(* IEC 61131-3 sources: Industry-PLC-LLM/data/PLCBEAD_repo/PLCBEAD_PLCEmbed-main/PLC-BEAD/Source/PLC_Programs (part 15) *)

(* ---- INC.ST ---- *)
FUNCTION INC:INT
	VAR_INPUT
		X :	INT;
		D :	INT;
		M :	INT;
	END_VAR

	inc := (X + D + M + 1) MOD (M + 1);
END_FUNCTION

PROGRAM program0
  VAR
    LocalVar0 : INT;
	LocalVar1 : INT;
	LocalVar2 : INT;
	LocalOUT  : INT;
  END_VAR
  	LocalOUT := INC(LocalVar0, LocalVar1,LocalVar2);
END_PROGRAM

CONFIGURATION Config0
  RESOURCE Res0 ON PLC
    TASK task0(INTERVAL := T#20ms,PRIORITY := 0);
    PROGRAM instance0 WITH task0 : program0;
  END_RESOURCE
END_CONFIGURATION

(* ---- INC1.ST ---- *)
FUNCTION INC1:INT

	VAR_INPUT
		X :	INT;
		N :	INT;
	END_VAR

	IF X >= N - 1 THEN
		INC1 := 0;
	ELSE
		INC1 := X + 1;
	END_IF;
END_FUNCTION

PROGRAM program0
  VAR
	X :	INT;
	N :	INT;
    CEIL5_OUT : INT;
  END_VAR

  CEIL5_OUT := INC1(X, N);
END_PROGRAM

CONFIGURATION Config0

  RESOURCE Res0 ON PLC
    TASK task0(INTERVAL := T#20ms,PRIORITY := 0);
    PROGRAM instance0 WITH task0 : program0;
  END_RESOURCE
END_CONFIGURATION

(* ---- INC2.ST ---- *)
FUNCTION INC2:INT

	VAR_INPUT
		X :	INT;
		D :	INT;
		L :	INT;
		U :	INT;
	END_VAR

	VAR
		tmp :	INT;
	END_VAR

	tmp := U - L + 1;
	INC2 := (X + D - L + tmp) MOD tmp + L;

END_FUNCTION

PROGRAM program0
	VAR
		X :	INT;
		D :	INT;
		L :	INT;
		U :	INT;
		CEIL5_OUT : INT;
	END_VAR

  	CEIL5_OUT := INC2(X, D, L, U);
END_PROGRAM

CONFIGURATION Config0

	RESOURCE Res0 ON PLC
		TASK task0(INTERVAL := T#20ms,PRIORITY := 0);
		PROGRAM instance0 WITH task0 : program0;
	END_RESOURCE

END_CONFIGURATION

(* ---- INI_PARSER_BUF_DEMO.ST ---- *)
PROGRAM INI_PARSER_BUF_DEMO

	VAR

	END_VAR

	VAR_EXTERNAL

	END_VAR

	VAR
		SMTP_SERVER :	STRING;
		SMTP_FROM :	STRING;
		STATION_NAME :	STRING;
		STATION_IP :	STRING;
	END_VAR

	VAR
		IPB :	INI_PARSER_BUF;
		FS :	FILE_SERVER;
		FSD :	oscat_FILE_SERVER_DATA;
		PT :	oscat_NETWORK_BUFFER;
		section :	INT;
		key :	oscat_STRING250;
		value :	oscat_STRING250;
		str :	oscat_STRING250;
		step :	INT;
		result :	BYTE;
		offset :	UDINT;
		run :	BYTE;
		done :	BOOL;
	END_VAR

	CASE step OF

	00:	IF NOT done then
			FSD.FILENAME := 'config.ini';
			FSD.MODE := BYTE#1;
			FSD.OFFSET := UDINT#0;
			FSD.AUTO_CLOSE := T#0s;
			PT.SIZE := UINT#65535;
			step := 10;
		END_IF;

	10:	IF FSD.MODE = BYTE#0 THEN
			offset := UDINT#0;
			str := '';
			run := BYTE#3;
			step := 50;
		END_IF;

	50:	IF run = BYTE#0 THEN
			run := BYTE#3;

			IF result = BYTE#1 THEN
				IF EQ_STRING(key,'Station') THEN
					section := 1;
				ELSIF EQ_STRING(key,'SMTP') THEN
					section := 2;

				ELSE
					section := 0;
				END_IF;

			ELSIF result = BYTE#2 AND section > 0 THEN

				CASE section OF

				1:
					IF EQ_STRING(key,'NAME') THEN
						STATION_NAME := value;
					ELSIF EQ_STRING(key,'IP') THEN
						STATION_IP := value;
					END_IF;

				2:
					IF EQ_STRING(key,'SERVER') THEN
						SMTP_SERVER := value;
					ELSIF EQ_STRING(key,'FROM') THEN
						SMTP_FROM := value;
					END_IF;

				END_CASE;

			ELSIF result = BYTE#10 THEN
				run := BYTE#0;
				FSD.MODE := BYTE#5;
				step := 80;
			END_IF;
		END_IF;

	80:	IF FSD.MODE = BYTE#0 THEN
			done := TRUE;
			step := 0;
		END_IF;

	END_CASE;

	IPB(STR:=str,RUN:=run,OFFSET:=offset,KEY:=key,VALUE:=value,PT:=PT);
	str:=IPB.STR;
	run:=IPB.RUN;
	offset:=IPB.OFFSET;
	key:=IPB.KEY;
	value:=IPB.VALUE;
	PT:=IPB.PT;
	result:=IPB.RESULT;

	FS(FSD:=FSD,PT:=PT);
	FSD:=FS.FSD;
	PT:=FS.PT;

END_PROGRAM

(* ---- INI_PARSER_FILE_DEMO.ST ---- *)
PROGRAM INI_PARSER_FILE_DEMO

	VAR

	END_VAR

	VAR_EXTERNAL

	END_VAR

	VAR
		SMTP_SERVER :	STRING;
		SMTP_FROM :	STRING;
		STATION_NAME :	STRING;
		STATION_IP :	STRING;
	END_VAR

	VAR
		IPF :	INI_PARSER_FILE;
		FS :	FILE_SERVER;
		FSD :	oscat_FILE_SERVER_DATA;
		PT :	oscat_NETWORK_BUFFER;
		section :	INT;
		filename :	STRING;
		key :	oscat_STRING250;
		value :	oscat_STRING250;
		str :	oscat_STRING250;
		step :	INT;
		result :	BYTE;
		offset :	UDINT;
		run :	BYTE;
		done :	BOOL;
	END_VAR

	CASE step OF

	00:	IF NOT done THEN
			filename := 'config.ini';
			offset := UDINT#0;
			str := '';
			run := BYTE#3;
			step := 50;
		END_IF;

	50:	IF run = BYTE#0 THEN

			run := BYTE#3;

			IF result = BYTE#1 THEN
				IF EQ_STRING(key,'Station') THEN
					section := 1;
				ELSIF EQ_STRING(key,'SMTP') THEN
					section := 2;

				ELSE
					section := 0;
				END_IF;

			ELSIF result = BYTE#2 AND section > 0 THEN

				CASE section OF

				1:
					IF EQ_STRING(key,'NAME') THEN
						STATION_NAME := value;
					ELSIF EQ_STRING(key,'IP') THEN
						STATION_IP := value;
					END_IF;

				2:
					IF EQ_STRING(key,'SERVER') THEN
						SMTP_SERVER := value;
					ELSIF EQ_STRING(key,'FROM') THEN
						SMTP_FROM := value;
					END_IF;

				END_CASE;

			ELSIF result = BYTE#10 THEN
				run := BYTE#0;
				FSD.MODE := BYTE#5;
				step := 30;
			END_IF;
		END_IF;

	30:	IF FSD.MODE = BYTE#0 THEN
			step := 0;
			done := TRUE;
		END_IF;

	END_CASE;

	IPF(FILENAME:=FILENAME,FSD:=FSD,STR:=str,RUN:=run,OFFSET:=offset,KEY:=key,VALUE:=value,PT:=PT);
	FILENAME:=IPF.FILENAME;
	FSD:=IPF.FSD;
	str:=IPF.STR;
	run:=IPF.RUN;
	offset:=IPF.OFFSET;
	key:=IPF.KEY;
	value:=IPF.VALUE;
	PT:=IPF.PT;
	result:=IPF.RESULT;

	FS(FSD:=FSD,PT:=PT);
	FSD:=FS.FSD;
	PT:=FS.PT;

END_PROGRAM

(* ---- INT_TO_BCDC.ST ---- *)
FUNCTION INT_TO_BCDC:BYTE

	VAR_INPUT
		IN :	INT;
	END_VAR

	INT_TO_BCDC := SHL(INT_TO_BYTE(IN / INT#10),4) OR INT_TO_BYTE(in MOD INT#10);

END_FUNCTION

PROGRAM program0

	VAR
		IN :	INT;
		OUT : BYTE;
	END_VAR

	OUT := INT_TO_BCDC(IN);

END_PROGRAM

CONFIGURATION Config0

	RESOURCE Res0 ON PLC
		TASK task0(INTERVAL := T#20ms,PRIORITY := 0);
		PROGRAM instance0 WITH task0 : program0;
	END_RESOURCE

END_CONFIGURATION

(* ---- INT_TO_TIME.ST ---- *)
FUNCTION _INT_TO_TIME:TIME

	VAR_INPUT
		IN :	INT;
	END_VAR

	_INT_TO_TIME := DINT_TO_TIME(INT_TO_DINT(IN));

END_FUNCTION

PROGRAM program0
	VAR
		IN :	INT;
		OUT : TIME;
	END_VAR

	OUT := _INT_TO_TIME(IN);
END_PROGRAM

CONFIGURATION Config0

	RESOURCE Res0 ON PLC
		TASK task0(INTERVAL := T#20ms,PRIORITY := 0);
		PROGRAM instance0 WITH task0 : program0;
	END_RESOURCE

END_CONFIGURATION

(* ---- INV.ST ---- *)
FUNCTION INV:REAL

	VAR_INPUT
		X :	REAL;
	END_VAR

	IF X <> 0.0 THEN INV := 1.0 / X; END_IF;

END_FUNCTION

PROGRAM program0
	VAR
		X :	REAL;
		OUT : REAL;
	END_VAR

	OUT := INV(X);
END_PROGRAM

CONFIGURATION Config0

	RESOURCE Res0 ON PLC
		TASK task0(INTERVAL := T#20ms,PRIORITY := 0);
		PROGRAM instance0 WITH task0 : program0;
	END_RESOURCE

END_CONFIGURATION

(* ---- IP4_CHECK.ST ---- *)
FUNCTION IP4_CHECK:BOOL

	VAR_INPUT
		NIP :	DWORD;
		LIP :	DWORD;
		SM :	DWORD;
	END_VAR

	IP4_CHECK := (NIP AND sm) = (LIP AND SM);

END_FUNCTION

PROGRAM program0
	VAR
		NIP :	DWORD;
		LIP :	DWORD;
		SM :	DWORD;
		CEIL5_OUT : BOOL;
	END_VAR

  	CEIL5_OUT := IP4_CHECK(NIP, LIP, SM);
END_PROGRAM

CONFIGURATION Config0

  RESOURCE Res0 ON PLC
    TASK task0(INTERVAL := T#20ms,PRIORITY := 0);
    PROGRAM instance0 WITH task0 : program0;
  END_RESOURCE
END_CONFIGURATION

(* ---- IS_URLCHR.ST ---- *)
FUNCTION IS_URLCHR:BOOL

	VAR_INPUT
		IN :	BYTE;
	END_VAR

	IS_URLCHR := ((IN>BYTE#47) AND (IN<BYTE#58)) OR ((IN>BYTE#64) AND (IN<BYTE#91)) OR ((IN>BYTE#96) AND (IN<BYTE#123)) OR (in=BYTE#126) OR (in=BYTE#95) OR (in=BYTE#45) OR (in=BYTE#46);

END_FUNCTION

PROGRAM program0
	VAR
		IN :	BYTE;
		CEIL5_OUT : BOOL;
	END_VAR

  	CEIL5_OUT := IS_URLCHR(IN);
END_PROGRAM

CONFIGURATION Config0

  RESOURCE Res0 ON PLC
    TASK task0(INTERVAL := T#20ms,PRIORITY := 0);
    PROGRAM instance0 WITH task0 : program0;
  END_RESOURCE
END_CONFIGURATION

(* ---- ISC_ALPHA.ST ---- *)
FUNCTION SETUP_EXTENDED_ASCII:BOOL

	VAR_INPUT
		X :	BOOL;
	END_VAR

	SETUP_EXTENDED_ASCII := X OR TRUE;

END_FUNCTION

FUNCTION ISC_ALPHA:BOOL

	VAR_INPUT
		IN :	BYTE;
	END_VAR

	IF SETUP_EXTENDED_ASCII(FALSE) THEN
		ISC_ALPHA := (in > BYTE#64 AND in < BYTE#91) OR (in > BYTE#191  AND in <> BYTE#215 AND in <> BYTE#247) OR (in > BYTE#96 AND in < BYTE#123);
	ELSE
		ISC_ALPHA := (IN > BYTE#64 AND IN < BYTE#91) OR (in > BYTE#96 AND in < BYTE#123);
	END_IF;

END_FUNCTION

PROGRAM program0
	VAR
		IN : BYTE;
		OUT : BOOL;
	END_VAR

	OUT := ISC_ALPHA(IN);
END_PROGRAM

CONFIGURATION Config0

	RESOURCE Res0 ON PLC
		TASK task0(INTERVAL := T#20ms,PRIORITY := 0);
		PROGRAM instance0 WITH task0 : program0;
	END_RESOURCE

END_CONFIGURATION

(* ---- ISC_CTRL.ST ---- *)
FUNCTION ISC_CTRL:BOOL

	VAR_INPUT
		IN :	BYTE;
	END_VAR

	ISC_CTRL := IN < BYTE#32 OR IN = BYTE#127;

END_FUNCTION

PROGRAM program0
	VAR
		IN : BYTE;
		OUT : BOOL;
	END_VAR

	OUT := ISC_CTRL(IN);
END_PROGRAM

CONFIGURATION Config0

	RESOURCE Res0 ON PLC
		TASK task0(INTERVAL := T#20ms,PRIORITY := 0);
		PROGRAM instance0 WITH task0 : program0;
	END_RESOURCE

END_CONFIGURATION

(* ---- ISC_HEX.ST ---- *)
FUNCTION ISC_HEX:BOOL

	VAR_INPUT
		IN :	BYTE;
	END_VAR

	ISC_HEX := (IN > BYTE#47 AND IN < BYTE#58) OR (IN > BYTE#64 AND IN < BYTE#71) OR (IN > BYTE#96 AND IN < BYTE#103);

END_FUNCTION

PROGRAM program0
	VAR
		IN : BYTE;
		OUT : BOOL;
	END_VAR

	OUT := ISC_HEX(IN);
END_PROGRAM

CONFIGURATION Config0

	RESOURCE Res0 ON PLC
		TASK task0(INTERVAL := T#20ms,PRIORITY := 0);
		PROGRAM instance0 WITH task0 : program0;
	END_RESOURCE

END_CONFIGURATION

(* ---- ISC_LOWER.ST ---- *)
FUNCTION SETUP_EXTENDED_ASCII:BOOL

	VAR_INPUT
		X :	BOOL;
	END_VAR

	SETUP_EXTENDED_ASCII := X OR TRUE;

END_FUNCTION

FUNCTION ISC_LOWER:BOOL

	VAR_INPUT
		IN :	BYTE;
	END_VAR

	IF SETUP_EXTENDED_ASCII(FALSE) THEN
		ISC_LOWER := ((in > BYTE#96) AND (in < BYTE#123)) OR ((in > BYTE#222) AND (in <> BYTE#247));
	ELSE
		ISC_LOWER := ((in > BYTE#96) AND (in < BYTE#123));
	END_IF;

END_FUNCTION

PROGRAM program0
	VAR
		IN : BYTE;
		OUT : BOOL;
	END_VAR

	OUT := ISC_LOWER(IN);
END_PROGRAM

CONFIGURATION Config0

	RESOURCE Res0 ON PLC
		TASK task0(INTERVAL := T#20ms,PRIORITY := 0);
		PROGRAM instance0 WITH task0 : program0;
	END_RESOURCE

END_CONFIGURATION

(* ---- ISC_NUM.ST ---- *)
FUNCTION ISC_NUM:BOOL

	VAR_INPUT
		IN :	BYTE;
	END_VAR

	ISC_NUM := IN > BYTE#47 AND IN < BYTE#58;

END_FUNCTION

PROGRAM program0
	VAR
		IN : BYTE;
		OUT : BOOL;
	END_VAR

	OUT := ISC_NUM(IN);
END_PROGRAM

CONFIGURATION Config0

	RESOURCE Res0 ON PLC
		TASK task0(INTERVAL := T#20ms,PRIORITY := 0);
		PROGRAM instance0 WITH task0 : program0;
	END_RESOURCE

END_CONFIGURATION

(* ---- ISC_UPPER.ST ---- *)
FUNCTION SETUP_EXTENDED_ASCII:BOOL

	VAR_INPUT
		X :	BOOL;
	END_VAR

	SETUP_EXTENDED_ASCII := X OR TRUE;

END_FUNCTION

FUNCTION ISC_UPPER:BOOL

	VAR_INPUT
		IN :	BYTE;
	END_VAR

	IF SETUP_EXTENDED_ASCII(FALSE) THEN
		ISC_UPPER :=  ((in > BYTE#64) AND (in < BYTE#91)) OR (((in > BYTE#191) AND (in < BYTE#223)) AND (in <> BYTE#215));
	ELSE
		ISC_UPPER := ((in > BYTE#64) AND (in < BYTE#91));
	END_IF;

END_FUNCTION

PROGRAM program0
	VAR
		IN : BYTE;
		OUT : BOOL;
	END_VAR

	OUT := ISC_UPPER(IN);
END_PROGRAM

CONFIGURATION Config0

	RESOURCE Res0 ON PLC
		TASK task0(INTERVAL := T#20ms,PRIORITY := 0);
		PROGRAM instance0 WITH task0 : program0;
	END_RESOURCE

END_CONFIGURATION

(* ---- JD2000.ST ---- *)
FUNCTION JD2000:REAL

	VAR_INPUT
		DTI :	UDINT;
	END_VAR

	JD2000 := UDINT_TO_REAL(DTI - UDINT#946728000) / 86400.0;

END_FUNCTION

PROGRAM program0
	VAR
		DTI :	UDINT;
		OUT : REAL;
	END_VAR

	OUT := JD2000(DTI);
END_PROGRAM

CONFIGURATION Config0

	RESOURCE Res0 ON PLC
		TASK task0(INTERVAL := T#20ms,PRIORITY := 0);
		PROGRAM instance0 WITH task0 : program0;
	END_RESOURCE

END_CONFIGURATION

(* ---- K_TO_C.ST ---- *)
FUNCTION K_TO_C:REAL

	VAR_INPUT
		KELVIN :	REAL;
	END_VAR

	K_to_C := Kelvin + 273.15;

END_FUNCTION

PROGRAM program0
	VAR
		KELVIN : REAL;
		OUT : REAL;
	END_VAR

	OUT := K_TO_C(KELVIN);
END_PROGRAM

CONFIGURATION Config0

	RESOURCE Res0 ON PLC
		TASK task0(INTERVAL := T#20ms,PRIORITY := 0);
		PROGRAM instance0 WITH task0 : program0;
	END_RESOURCE

END_CONFIGURATION

(* ---- KMH_TO_MS.ST ---- *)
FUNCTION KMH_TO_MS:REAL

	VAR_INPUT
		KMH :	REAL;
	END_VAR

	KMH_TO_MS := kmh * 0.2777777777777;

END_FUNCTION

PROGRAM program0
	VAR
		KMH : REAL;
		OUT : REAL;
	END_VAR

	OUT := KMH_TO_MS(KMH);
END_PROGRAM

CONFIGURATION Config0

	RESOURCE Res0 ON PLC
		TASK task0(INTERVAL := T#20ms,PRIORITY := 0);
		PROGRAM instance0 WITH task0 : program0;
	END_RESOURCE

END_CONFIGURATION

(* ---- LANGEVIN.ST ---- *)
FUNCTION COTH:REAL

	VAR_INPUT
		X :	REAL;
	END_VAR

	IF X > 20.0 THEN
		COTH :=1.0;
	ELSIF X < -20.0 THEN
		COTH := -1.0;
	ELSE
		COTH := 1.0 + 2.0 / (EXP(X * 2.0) - 1.0);
	END_IF;

END_FUNCTION

FUNCTION LANGEVIN:REAL

	VAR_INPUT
		X :	REAL;
	END_VAR

	IF X = 0.0 THEN
		LANGEVIN := 0.0;
	ELSE
		LANGEVIN := COTH(X) - 1.0 / X;
	END_IF;

END_FUNCTION

PROGRAM program0
	VAR
		X :	REAL;
		OUT : REAL;
	END_VAR

	OUT := LANGEVIN(X);
END_PROGRAM

CONFIGURATION Config0

	RESOURCE Res0 ON PLC
		TASK task0(INTERVAL := T#20ms,PRIORITY := 0);
		PROGRAM instance0 WITH task0 : program0;
	END_RESOURCE

END_CONFIGURATION

(* ---- LEAP_DAY.ST ---- *)
FUNCTION LEAP_DAY:BOOL

	VAR_INPUT
		IDATE :	UDINT;
	END_VAR

	LEAP_DAY := IDATE MOD UDINT#126230400 = UDINT#68169600;

END_FUNCTION

PROGRAM program0
	VAR
		IDATE :	UDINT;
		OUT : BOOL;
	END_VAR

	OUT := LEAP_DAY(IDATE);
END_PROGRAM

CONFIGURATION Config0

	RESOURCE Res0 ON PLC
		TASK task0(INTERVAL := T#20ms,PRIORITY := 0);
		PROGRAM instance0 WITH task0 : program0;
	END_RESOURCE

END_CONFIGURATION

(* ---- LEAP_OF_DATE.ST ---- *)
FUNCTION LEAP_OF_DATE:BOOL

	VAR_INPUT
		IDATE :	UDINT;
	END_VAR

	LEAP_OF_DATE := SHL(UDINT_TO_DWORD((idate + UDINT#43200) / UDINT#31557600), 30) = DWORD#16#80000000;

END_FUNCTION

PROGRAM program0
  VAR
    LocalVar0 : UDINT;
	LocalOUT  : BOOL;
  END_VAR
  	LocalOUT := LEAP_OF_DATE(LocalVar0);
END_PROGRAM

CONFIGURATION Config0
  RESOURCE Res0 ON PLC
    TASK task0(INTERVAL := T#20ms,PRIORITY := 0);
    PROGRAM instance0 WITH task0 : program0;
  END_RESOURCE
END_CONFIGURATION

(* ---- LEAP_YEAR.ST ---- *)
FUNCTION LEAP_YEAR:BOOL

  VAR_INPUT
    YEAR :	INT;
  END_VAR

  IF (year MOD INT#400) = INT#00 THEN
    leap_year := TRUE;
  ELSIF (year MOD INT#100) = INT#00 THEN
    leap_year := FALSE;
  ELSIF (year MOD INT#04) = INT#00 THEN
    leap_year := TRUE;
  ELSE
    leap_year := FALSE;
  END_IF;

END_FUNCTION

PROGRAM program0
	VAR
		YEAR :	INT;
		OUT : BOOL;
	END_VAR

	OUT := LEAP_YEAR(YEAR);
END_PROGRAM

CONFIGURATION Config0

	RESOURCE Res0 ON PLC
		TASK task0(INTERVAL := T#20ms,PRIORITY := 0);
		PROGRAM instance0 WITH task0 : program0;
	END_RESOURCE

END_CONFIGURATION

(* ---- LTIME_TO_UTC.ST ---- *)
FUNCTION _INT_TO_UDINT:UDINT
	VAR_INPUT
		IN :	INT;
	END_VAR

	_INT_TO_UDINT := DINT_TO_UDINT(INT_TO_DINT(IN));
END_FUNCTION

FUNCTION LTIME_TO_UTC:UDINT

	VAR_INPUT
		LTIME :	UDINT;
		DST :	BOOL;
		TIME_ZONE_OFFSET :	INT;
	END_VAR

	LTIME_TO_UTC := LTIME - _INT_TO_UDINT(TIME_ZONE_OFFSET * 60);
	IF DST THEN LTIME_TO_UTC := LTIME_TO_UTC - UDINT#3600; END_IF;

END_FUNCTION

PROGRAM program0
	VAR
		LTIME :	UDINT;
		DST :	BOOL;
		TIME_ZONE_OFFSET :	INT;
		CEIL5_OUT : UDINT;
	END_VAR

  CEIL5_OUT := LTIME_TO_UTC(LTIME, DST, TIME_ZONE_OFFSET);
END_PROGRAM

CONFIGURATION Config0

  RESOURCE Res0 ON PLC
    TASK task0(INTERVAL := T#20ms,PRIORITY := 0);
    PROGRAM instance0 WITH task0 : program0;
  END_RESOURCE
END_CONFIGURATION

(* ---- MANUAL.ST ---- *)
FUNCTION MANUAL:BOOL

	VAR_INPUT
		_IN :	BOOL;
		_ON :	BOOL;
		OFF :	BOOL;
	END_VAR

	MANUAL := NOT OFF AND (_IN OR _ON);

END_FUNCTION

PROGRAM program0
	VAR
		_IN :	BOOL;
		_ON :	BOOL;
		OFF :	BOOL;

		OUT : BOOL;
	END_VAR

	OUT := MANUAL(_IN, _ON, OFF);

END_PROGRAM

CONFIGURATION Config0

	RESOURCE Res0 ON PLC
		TASK task0(INTERVAL := T#20ms,PRIORITY := 0);
		PROGRAM instance0 WITH task0 : program0;
	END_RESOURCE

END_CONFIGURATION

(* ---- MAX3.ST ---- *)
FUNCTION MAX3:REAL

	VAR_INPUT
		IN1 :	REAL;
		IN2 :	REAL;
		IN3 :	REAL;
	END_VAR

	MAX3 := MAX(MAX(IN1,IN2),IN3);

END_FUNCTION

PROGRAM program0
	VAR
		IN1 :	REAL;
		IN2 :	REAL;
		IN3 :	REAL;

		OUT : REAL;
	END_VAR

	OUT := MAX3(IN1, IN2, IN3);

END_PROGRAM

CONFIGURATION Config0

	RESOURCE Res0 ON PLC
		TASK task0(INTERVAL := T#20ms,PRIORITY := 0);
		PROGRAM instance0 WITH task0 : program0;
	END_RESOURCE

END_CONFIGURATION

(* ---- MAX_TIME.ST ---- *)
FUNCTION _MAX_TIME:TIME

	VAR_INPUT
		IN1 :	TIME;
		IN2 :	TIME;
	END_VAR

	_MAX_TIME := SEL_TIME(IN1 < IN2,IN1,IN2);

END_FUNCTION

PROGRAM program0
	VAR
		IN1 :	TIME;
		IN2 :	TIME;

		OUT : TIME;
	END_VAR

	OUT := _MAX_TIME(IN1, IN2);

END_PROGRAM

CONFIGURATION Config0

	RESOURCE Res0 ON PLC
		TASK task0(INTERVAL := T#20ms,PRIORITY := 0);
		PROGRAM instance0 WITH task0 : program0;
	END_RESOURCE

END_CONFIGURATION

(* ---- MD5_AUX.ST ---- *)
FUNCTION MD5_AUX:DWORD

	VAR_INPUT
		N :	INT;
		A :	DWORD;
		B :	DWORD;
		C :	DWORD;
		D :	DWORD;
		X :	DWORD;
		U :	INT;
		T :	DWORD;
	END_VAR

	VAR
		w :	DWORD;
	END_VAR

	CASE N OF
		1: w := (B AND C) OR (NOT(B) AND D);
		2: w := (B AND D) OR (C AND NOT D);
		3: w := (B XOR C XOR D);
		4: w := (C XOR (B OR  NOT(D)));
	END_CASE;

	MD5_AUX := UDINT_TO_DWORD(DWORD_TO_UDINT(B) + DWORD_TO_UDINT(ROL_DWORD(UDINT_TO_DWORD(DWORD_TO_UDINT(A) + DWORD_TO_UDINT(w) + DWORD_TO_UDINT(X) + DWORD_TO_UDINT(T)),U)));

END_FUNCTION

PROGRAM program0
	VAR
		N :	INT;
		A :	DWORD;
		B :	DWORD;
		C :	DWORD;
		D :	DWORD;
		X :	DWORD;
		U :	INT;
		T :	DWORD;
		CEIL5_OUT : DWORD;
	END_VAR

  	CEIL5_OUT := MD5_AUX(N, A, B, C, D, X, U, T);
END_PROGRAM

CONFIGURATION Config0

  RESOURCE Res0 ON PLC
    TASK task0(INTERVAL := T#20ms,PRIORITY := 0);
    PROGRAM instance0 WITH task0 : program0;
  END_RESOURCE
END_CONFIGURATION

(* ---- MID3.ST ---- *)
FUNCTION MID3:REAL

	VAR_INPUT
		IN1 :	REAL;
		IN2 :	REAL;
		IN3 :	REAL;
	END_VAR

	VAR
		_IN1 :	REAL;
		_IN2 :	REAL;
		_IN3 :	REAL;
	END_VAR

	_IN1 := IN1;
	_IN2 := IN2;
	_IN3 := IN3;

	IF _IN1 > _IN2 THEN MID3 := _IN1; _IN1 := _IN2; _IN2 := MID3; END_IF;
	IF _IN2 > _IN3 THEN _IN2 := _IN3; END_IF;
	MID3 := SEL(_IN1 > _IN2, _IN2, _IN1);

END_FUNCTION

PROGRAM program0
	VAR
		IN1 :	REAL;
		IN2 :	REAL;
		IN3 :	REAL;

		OUT : REAL;
	END_VAR

	OUT := MID3(IN1, IN2, IN3);

END_PROGRAM

CONFIGURATION Config0

	RESOURCE Res0 ON PLC
		TASK task0(INTERVAL := T#20ms,PRIORITY := 0);
		PROGRAM instance0 WITH task0 : program0;
	END_RESOURCE

END_CONFIGURATION

(* ---- MIN3.ST ---- *)
FUNCTION MIN3:REAL

	VAR_INPUT
		IN1 :	REAL;
		IN2 :	REAL;
		IN3 :	REAL;
	END_VAR

	MIN3 := MIN(MIN(IN1,IN2),IN3);

END_FUNCTION

PROGRAM program0

	VAR
		IN1 :	REAL;
		IN2 :	REAL;
		IN3 :	REAL;
		CEIL5_OUT : REAL;
	END_VAR

	CEIL5_OUT := MIN3(IN1, IN2, IN3);

END_PROGRAM

CONFIGURATION Config0

	RESOURCE Res0 ON PLC
		TASK task0(INTERVAL := T#20ms,PRIORITY := 0);
		PROGRAM instance0 WITH task0 : program0;
	END_RESOURCE

END_CONFIGURATION

(* ---- MINUTE.ST ---- *)
FUNCTION MINUTE:INT

	VAR_INPUT
		ITOD :	UDINT;
	END_VAR

	minute := UDINT_TO_INT((itod / UDINT#60000) - ((itod / UDINT#3600000) * UDINT#60));

END_FUNCTION

PROGRAM program0
  VAR
	  ITOD :	UDINT;
    CEIL5_OUT : INT;
  END_VAR

  CEIL5_OUT := MINUTE(ITOD);
END_PROGRAM

CONFIGURATION Config0

  RESOURCE Res0 ON PLC
    TASK task0(INTERVAL := T#20ms,PRIORITY := 0);
    PROGRAM instance0 WITH task0 : program0;
  END_RESOURCE
END_CONFIGURATION

(* ---- MINUTE_OF_DT.ST ---- *)
FUNCTION MINUTE_OF_DT:INT
	VAR_INPUT
		XDT :	UDINT;
	END_VAR

	MINUTE_OF_DT := UDINT_TO_INT((XDT MOD UDINT#3600) / UDINT#60);
END_FUNCTION

PROGRAM program0
  VAR
    LocalVar0 : UDINT;
	LocalOUT  : INT;
  END_VAR
  	LocalOUT := MINUTE_OF_DT(LocalVar0);
END_PROGRAM

CONFIGURATION Config0
  RESOURCE Res0 ON PLC
    TASK task0(INTERVAL := T#20ms,PRIORITY := 0);
    PROGRAM instance0 WITH task0 : program0;
  END_RESOURCE
END_CONFIGURATION

(* ---- MINUTE_TO_TIME.ST ---- *)
FUNCTION _REAL_TO_UDINT:UDINT

  	VAR_INPUT
		X :	REAL;
	END_VAR

	IF REAL_TO_UDINT(0.5) = UDINT#1 THEN
		_REAL_TO_UDINT := REAL_TO_UDINT(x);
	ELSIF X > 0.0 THEN
		_REAL_TO_UDINT := REAL_TO_UDINT(x+0.5);
	ELSIF X < 0.0 THEN
		_REAL_TO_UDINT := REAL_TO_UDINT(x-0.5);
	ELSE
		_REAL_TO_UDINT := UDINT#0;
	END_IF;

END_FUNCTION

FUNCTION MINUTE_TO_TIME:TIME

	VAR_INPUT
		IN :	REAL;
	END_VAR

	minute_to_time := UDINT_TO_TIME(_REAL_TO_UDINT(IN * 60000.0));

END_FUNCTION

PROGRAM program0

	VAR
		IN :	REAL;
		CEIL5_OUT : TIME;
	END_VAR

	CEIL5_OUT := MINUTE_TO_TIME(IN);

END_PROGRAM

CONFIGURATION Config0

	RESOURCE Res0 ON PLC
		TASK task0(INTERVAL := T#20ms,PRIORITY := 0);
		PROGRAM instance0 WITH task0 : program0;
	END_RESOURCE

END_CONFIGURATION

(* ---- MIX.ST ---- *)
FUNCTION MIX:REAL

	VAR_INPUT
		A :	REAL;
		B :	REAL;
		M :	REAL;
	END_VAR

	MIX := (1.0 - M) * A + M * B;

END_FUNCTION

PROGRAM program0
	VAR
		A :	REAL;
		B :	REAL;
		M :	REAL;

		OUT : REAL;
	END_VAR

	OUT := MIX(A, B, M);

END_PROGRAM

CONFIGURATION Config0

	RESOURCE Res0 ON PLC
		TASK task0(INTERVAL := T#20ms,PRIORITY := 0);
		PROGRAM instance0 WITH task0 : program0;
	END_RESOURCE

END_CONFIGURATION

(* ---- MODR.ST ---- *)
FUNCTION FLOOR2 : DINT
	VAR_INPUT
		x : REAL;
	END_VAR

	FLOOR2 := REAL_TO_DINT(X);
	IF DINT_TO_REAL(FLOOR2) > X THEN
		FLOOR2 := FLOOR2 - DINT#1;
	END_IF;

END_FUNCTION

FUNCTION MODR: REAL

	VAR_INPUT
		IN :	REAL;
		DIVI :	REAL;
	END_VAR

	IF divi = 0.0 THEN
		MODR := 0.0;
	ELSE
		MODR := in - DINT_TO_REAL(FLOOR2(in / divi)) * divi;
	END_IF;

END_FUNCTION

PROGRAM program0

  	VAR
		IN :	REAL;
		DIVI :	REAL;
		CEIL5_OUT : REAL;
  	END_VAR

  	CEIL5_OUT := MODR(IN, DIVI);
END_PROGRAM

CONFIGURATION Config0

  RESOURCE Res0 ON PLC
    TASK task0(INTERVAL := T#20ms,PRIORITY := 0);
    PROGRAM instance0 WITH task0 : program0;
  END_RESOURCE
END_CONFIGURATION

(* ---- MONTH_BEGIN.ST ---- *)
FUNCTION LEAP_OF_DATE:BOOL

	VAR_INPUT
		IDATE :	UDINT;
	END_VAR

	LEAP_OF_DATE := SHL(UDINT_TO_DWORD((idate + UDINT#43200) / UDINT#31557600), 30) = DWORD#16#80000000;
END_FUNCTION

FUNCTION DAY_OF_YEAR:INT
	VAR_INPUT
		IDATE :	UDINT;
	END_VAR

	DAY_OF_YEAR := UDINT_TO_INT(((idate) / UDINT#86400) MOD UDINT#1461);
	IF DAY_OF_YEAR > 729 THEN
		IF DAY_OF_YEAR > 1095 THEN DAY_OF_YEAR := DAY_OF_YEAR - 1095; ELSE DAY_OF_YEAR := DAY_OF_YEAR - 729; END_IF;
	ELSIF DAY_OF_YEAR > 364 THEN
		DAY_OF_YEAR := DAY_OF_YEAR - 364;
	ELSE
		DAY_OF_YEAR := DAY_OF_YEAR + 1;
	END_IF;
END_FUNCTION

FUNCTION MONTH_OF_DATE:INT

	VAR_INPUT
		IDATE :	UDINT;
	END_VAR

	MONTH_OF_DATE := DAY_OF_YEAR(idate);
	IF MONTH_OF_DATE < 32 THEN
		MONTH_OF_DATE := 1;
	ELSIF LEAP_OF_DATE((IDATE)) THEN
		MONTH_OF_DATE := (MONTH_OF_DATE * 53 + 1668) / 1623;
	ELSE
		MONTH_OF_DATE := (MONTH_OF_DATE * 53 + 1700) / 1620;
	END_IF;
END_FUNCTION

FUNCTION DAY_OF_MONTH:INT
	VAR_INPUT
		IDATE :	UDINT;
	END_VAR

	day_of_month := day_of_year(idate);

	IF leap_of_Date((idate)) THEN
		CASE day_of_month OF
			32..60	:	day_of_month := day_of_month - 31;
			61..91	:	day_of_month := day_of_month - 60;
			92..121 :	day_of_month := day_of_month - 91;
			122..152:	day_of_month := day_of_month - 121;
			153..182:	day_of_month := day_of_month - 152;
			183..213:	day_of_month := day_of_month - 182;
			214..244:	day_of_month := day_of_month - 213;
			245..274:	day_of_month := day_of_month - 244;
			275..305:	day_of_month := day_of_month - 274;
			306..335:	day_of_month := day_of_month - 305;
			336..366:	day_of_month := day_of_month - 335;
		END_CASE;
	ELSE
		CASE day_of_month OF
			32..59	:	day_of_month := day_of_month - 31;
			60..90	:	day_of_month := day_of_month - 59;
			91..120 :	day_of_month := day_of_month - 90;
			121..151:	day_of_month := day_of_month - 120;
			152..181:	day_of_month := day_of_month - 151;
			182..212:	day_of_month := day_of_month - 181;
			213..243:	day_of_month := day_of_month - 212;
			244..273:	day_of_month := day_of_month - 243;
			274..304:	day_of_month := day_of_month - 273;
			305..334:	day_of_month := day_of_month - 304;
			335..365:	day_of_month := day_of_month - 334;
		END_CASE;
	END_IF;
END_FUNCTION

FUNCTION _INT_TO_UDINT:UDINT
	VAR_INPUT
		IN :	INT;
	END_VAR

	_INT_TO_UDINT := DINT_TO_UDINT(INT_TO_DINT(IN));
END_FUNCTION

FUNCTION MONTH_BEGIN:UDINT

VAR_INPUT
	IDATE :	UDINT;
END_VAR

MONTH_BEGIN := idate - _INT_TO_UDINT(DAY_OF_MONTH(idate) - 1) * UDINT#86400;

END_FUNCTION

PROGRAM program0
	VAR
		IDATE :	UDINT;

		OUT : UDINT;
	END_VAR

	OUT := MONTH_BEGIN(IDATE);

END_PROGRAM

CONFIGURATION Config0

	RESOURCE Res0 ON PLC
		TASK task0(INTERVAL := T#20ms,PRIORITY := 0);
		PROGRAM instance0 WITH task0 : program0;
	END_RESOURCE

END_CONFIGURATION

(* ---- MONTH_END.ST ---- *)
FUNCTION LEAP_OF_DATE:BOOL

	VAR_INPUT
		IDATE :	UDINT;
	END_VAR

	LEAP_OF_DATE := SHL(UDINT_TO_DWORD((idate + UDINT#43200) / UDINT#31557600), 30) = DWORD#16#80000000;
END_FUNCTION

FUNCTION DAY_OF_YEAR:INT
	VAR_INPUT
		IDATE :	UDINT;
	END_VAR

	DAY_OF_YEAR := UDINT_TO_INT(((idate) / UDINT#86400) MOD UDINT#1461);
	IF DAY_OF_YEAR > 729 THEN
		IF DAY_OF_YEAR > 1095 THEN DAY_OF_YEAR := DAY_OF_YEAR - 1095; ELSE DAY_OF_YEAR := DAY_OF_YEAR - 729; END_IF;
	ELSIF DAY_OF_YEAR > 364 THEN
		DAY_OF_YEAR := DAY_OF_YEAR - 364;
	ELSE
		DAY_OF_YEAR := DAY_OF_YEAR + 1;
	END_IF;
END_FUNCTION

FUNCTION MONTH_OF_DATE:INT

	VAR_INPUT
		IDATE :	UDINT;
	END_VAR

	MONTH_OF_DATE := DAY_OF_YEAR(idate);
	IF MONTH_OF_DATE < 32 THEN
		MONTH_OF_DATE := 1;
	ELSIF LEAP_OF_DATE((IDATE)) THEN
		MONTH_OF_DATE := (MONTH_OF_DATE * 53 + 1668) / 1623;
	ELSE
		MONTH_OF_DATE := (MONTH_OF_DATE * 53 + 1700) / 1620;
	END_IF;
END_FUNCTION

FUNCTION YEAR_OF_DATE:INT
	VAR_INPUT
		IDATE :	UDINT;
	END_VAR

	YEAR_OF_DATE := UDINT_TO_INT((idate+UDINT#43200) / UDINT#31557600 + UDINT#1970);
END_FUNCTION

FUNCTION _INT_TO_UDINT:UDINT
	VAR_INPUT
		IN :	INT;
	END_VAR

	_INT_TO_UDINT := DINT_TO_UDINT(INT_TO_DINT(IN));
END_FUNCTION

FUNCTION DT_TO_DATE:UDINT
	VAR_INPUT
		IN :	UDINT;
	END_VAR

	DT_TO_DATE := (IN / UDINT#86400) * UDINT#86400;
END_FUNCTION

FUNCTION SET_DT:UDINT

	VAR_INPUT
		YEAR : INT;
		MONTH :	INT;
		DAY : INT;
		HOUR : INT;
		MINUTE : INT;
		SECOND : INT;
	END_VAR

	SET_DT := SET_DATE(YEAR, MONTH, DAY) + _INT_TO_UDINT(SECOND) + _INT_TO_UDINT(MINUTE) * UDINT#60 + _INT_TO_UDINT(HOUR) * UDINT#3600;

END_FUNCTION

FUNCTION SET_DATE:UDINT

	VAR_INPUT
		YEAR :	INT;
		MONTH :	INT;
		DAY :	INT;
	END_VAR

	VAR
		count :	INT;
	END_VAR

	IF month > 2 THEN
		count := (month - 1) * 30;
		IF month > 7 THEN
			count := count + DWORD_TO_INT(SHR(DINT_TO_DWORD(INT_TO_DINT(month) - INT_TO_DINT(3)),1));
		ELSE
			count := count + DWORD_TO_INT(SHR(DINT_TO_DWORD(INT_TO_DINT(month) - INT_TO_DINT(4)),1));
		END_IF;
		IF SHL(INT_TO_WORD(year),14) = WORD#0 THEN
			count := count + 1;
		END_IF;
	ELSE
		count := (month - 1) * 31;
	END_IF;
	SET_DATE := (_INT_TO_UDINT(count + day - 1) + DWORD_TO_UDINT(SHR(UDINT_TO_DWORD(_INT_TO_UDINT(year) * UDINT#1461 - UDINT#2878169), 2))) * UDINT#86400;

END_FUNCTION

FUNCTION MONTH_END:UDINT

	VAR_INPUT
		IDATE :	UDINT;
	END_VAR

	MONTH_END := SET_DATE(YEAR_OF_DATE(idate),MONTH_OF_DATE(idate)+1,1) - UDINT#86400;

END_FUNCTION

PROGRAM program0
	VAR
		IDATE :	UDINT;

		OUT : UDINT;
	END_VAR

	OUT := MONTH_END(IDATE);

END_PROGRAM

CONFIGURATION Config0

	RESOURCE Res0 ON PLC
		TASK task0(INTERVAL := T#20ms,PRIORITY := 0);
		PROGRAM instance0 WITH task0 : program0;
	END_RESOURCE

END_CONFIGURATION

(* ---- MONTH_OF_DATE.ST ---- *)
FUNCTION LEAP_OF_DATE:BOOL

	VAR_INPUT
		IDATE :	UDINT;
	END_VAR

	LEAP_OF_DATE := SHL(UDINT_TO_DWORD((idate + UDINT#43200) / UDINT#31557600), 30) = DWORD#16#80000000;

END_FUNCTION

FUNCTION DAY_OF_YEAR:INT
	VAR_INPUT
		IDATE :	DATE;
	END_VAR

	DAY_OF_YEAR := UDINT_TO_INT((DATE_TO_UDINT(idate) / UDINT#86400) MOD UDINT#1461);
	IF DAY_OF_YEAR > 729 THEN
		IF DAY_OF_YEAR > 1095 THEN DAY_OF_YEAR := DAY_OF_YEAR - 1095; ELSE DAY_OF_YEAR := DAY_OF_YEAR - 729; END_IF;
	ELSIF DAY_OF_YEAR > 364 THEN
		DAY_OF_YEAR := DAY_OF_YEAR - 364;
	ELSE
		DAY_OF_YEAR := DAY_OF_YEAR + 1;
	END_IF;
END_FUNCTION

FUNCTION MONTH_OF_DATE:INT

	VAR_INPUT
		IDATE :	DATE;
	END_VAR

	MONTH_OF_DATE := DAY_OF_YEAR(idate);
	IF MONTH_OF_DATE < 32 THEN
		MONTH_OF_DATE := 1;
	ELSIF LEAP_OF_DATE(DATE_TO_UDINT(IDATE)) THEN
		MONTH_OF_DATE := (MONTH_OF_DATE * 53 + 1668) / 1623;
	ELSE
		MONTH_OF_DATE := (MONTH_OF_DATE * 53 + 1700) / 1620;
	END_IF;

END_FUNCTION

PROGRAM program0
  VAR
    LocalVar0 : DATE;
	LocalOUT  : INT;
  END_VAR
  	LocalOUT := MONTH_OF_DATE(LocalVar0);
END_PROGRAM

CONFIGURATION Config0
  RESOURCE Res0 ON PLC
    TASK task0(INTERVAL := T#20ms,PRIORITY := 0);
    PROGRAM instance0 WITH task0 : program0;
  END_RESOURCE
END_CONFIGURATION

(* ---- MS_TO_BFT.ST ---- *)
FUNCTION MS_TO_BFT:INT

	VAR_INPUT
		MS :	REAL;
	END_VAR

	MS_TO_BFT := REAL_TO_INT(EXPT(MS * 1.196172, 0.666667));

END_FUNCTION

PROGRAM program0
	VAR
		MS :	REAL;

		OUT : INT;
	END_VAR

	OUT := MS_TO_BFT(MS);

END_PROGRAM

CONFIGURATION Config0

	RESOURCE Res0 ON PLC
		TASK task0(INTERVAL := T#20ms,PRIORITY := 0);
		PROGRAM instance0 WITH task0 : program0;
	END_RESOURCE

END_CONFIGURATION

(* ---- MS_TO_KMH.ST ---- *)
FUNCTION MS_TO_KMH:REAL

	VAR_INPUT
		MS :	REAL;
	END_VAR

	MS_TO_KMH := ms * 3.6;

END_FUNCTION

PROGRAM program0
	VAR
		MS :	REAL;

		OUT : REAL;
	END_VAR

	OUT := MS_TO_KMH(MS);

END_PROGRAM

CONFIGURATION Config0

	RESOURCE Res0 ON PLC
		TASK task0(INTERVAL := T#20ms,PRIORITY := 0);
		PROGRAM instance0 WITH task0 : program0;
	END_RESOURCE

END_CONFIGURATION

(* ---- MUL_ADD.ST ---- *)
FUNCTION MUL_ADD:REAL

	VAR_INPUT
		X :	REAL;
		K :	REAL;
		O :	REAL;
	END_VAR

	MUL_ADD := X * K + O;

END_FUNCTION

PROGRAM program0
	VAR
		X :	REAL;
		K :	REAL;
		O :	REAL;

		OUT : REAL;
	END_VAR

	OUT := MUL_ADD(X, K, O);

END_PROGRAM

CONFIGURATION Config0

	RESOURCE Res0 ON PLC
		TASK task0(INTERVAL := T#20ms,PRIORITY := 0);
		PROGRAM instance0 WITH task0 : program0;
	END_RESOURCE

END_CONFIGURATION

(* ---- MULTI_IN.ST ---- *)
FUNCTION MID3:REAL

	VAR_INPUT
		IN1 :	REAL;
		IN2 :	REAL;
		IN3 :	REAL;
	END_VAR

	VAR
		_IN1 :	REAL;
		_IN2 :	REAL;
		_IN3 :	REAL;
	END_VAR

	_IN1 := IN1;
	_IN2 := IN2;
	_IN3 := IN3;

	IF _IN1 > _IN2 THEN MID3 := _IN1; _IN1 := _IN2; _IN2 := MID3; END_IF;
	IF _IN2 > _IN3 THEN _IN2 := _IN3; END_IF;
	MID3 := SEL(_IN1 > _IN2, _IN2, _IN1);

END_FUNCTION

FUNCTION _BYTE_TO_INT:INT
	VAR_INPUT
		IN :	BYTE;
	END_VAR

	_BYTE_TO_INT := USINT_TO_INT(BYTE_TO_USINT(IN));
END_FUNCTION

FUNCTION MULTI_IN:REAL

	VAR_INPUT
		IN_1 :	REAL;
		IN_2 :	REAL;
		IN_3 :	REAL;
		DEFAULT :	REAL;
		IN_MIN :	REAL;
		IN_MAX :	REAL;
		MODE :	BYTE;
	END_VAR

	VAR
		count :	INT;
		F1 :	BOOL;
		F2 :	BOOL;
		F3 :	BOOL;
	END_VAR

	F1 :=  in_1 > in_min AND in_1 < in_max;
	F2 :=  in_2 > in_min AND in_2 < in_max;
	F3 :=  in_3 > in_min AND in_3 < in_max;

	CASE _BYTE_TO_INT(mode) OF
	0:	count := 0;
		IF F1 THEN
			count := count + 1;
			MULTI_IN := in_1;
		ELSE
			MULTI_IN := 0.0;
		END_IF;
		IF F2 THEN
			count := count + 1;
			MULTI_IN := MULTI_IN + in_2;
		END_IF;
		IF F3 THEN
			count := count + 1;
			MULTI_IN := MULTI_IN + in_3;
		END_IF;
		MULTI_IN := SEL_REAL(count = 0, MULTI_IN / INT_TO_REAL(count), default);

	1:	MULTI_IN := SEL_REAL(F1, default, IN_1);

	2:	MULTI_IN := SEL_REAL(F2, default, IN_2);

	3:	MULTI_IN := SEL_REAL(F3, default, IN_3);

	4:	MULTI_IN := default;

	5:	MULTI_IN := SEL_REAL(F1, in_max, IN_1);
		IF F2 AND in_2 < MULTI_IN THEN MULTI_IN := in_2; END_IF;
		IF F3 AND in_3 < MULTI_IN THEN MULTI_IN := in_3; END_IF;
		IF MULTI_IN = in_max THEN MULTI_IN := default; END_IF;

	6:	MULTI_IN := SEL_REAL(F1, in_min, IN_1);
		IF F2 AND in_2 > MULTI_IN THEN MULTI_IN := in_2; END_IF;
		IF F3 AND in_3 > MULTI_IN THEN MULTI_IN := in_3; END_IF;
		IF MULTI_IN = in_min THEN MULTI_IN := default; END_IF;

	7:	IF F1 AND F2 AND F3 THEN MULTI_IN := MID3(in_1, in_2, in_3);
		ELSIF F1 AND F2 THEN MULTI_IN := MIN(in_1, in_2);
		ELSIF F1 AND F3 THEN MULTI_IN := MIN(in_1, in_3);
		ELSIF F2 AND F3 THEN MULTI_IN := MIN(in_2, in_3);
		ELSIF F1 THEN MULTI_IN := in_1;
		ELSIF F2 THEN MULTI_IN := in_2;
		ELSIF F3 THEN MULTI_IN := in_3;
		ELSE MULTI_IN := default;
		END_IF;

	END_CASE;

END_FUNCTION

PROGRAM program0
	VAR
		IN_1 :	REAL;
		IN_2 :	REAL;
		IN_3 :	REAL;
		DEFAULT :	REAL;
		IN_MIN :	REAL;
		IN_MAX :	REAL;
		MODE :	BYTE;

		OUT : REAL;
	END_VAR

	OUT := MULTI_IN(IN_1, IN_2, IN_3, DEFAULT, IN_MIN, IN_MAX, MODE);

END_PROGRAM

CONFIGURATION Config0

	RESOURCE Res0 ON PLC
		TASK task0(INTERVAL := T#20ms,PRIORITY := 0);
		PROGRAM instance0 WITH task0 : program0;
	END_RESOURCE

END_CONFIGURATION

(* ---- MULTIME.ST ---- *)
FUNCTION _REAL_TO_DWORD: DWORD

  VAR_INPUT
    X :	REAL;
  END_VAR

  IF REAL_TO_DWORD(0.5) = DWORD#1 THEN
    _REAL_TO_DWORD := REAL_TO_DWORD(x);
  ELSIF X > 0.0 THEN
    _REAL_TO_DWORD := REAL_TO_DWORD(x+0.5);
  ELSIF X < 0.0 THEN
    _REAL_TO_DWORD := REAL_TO_DWORD(x-0.5);
  ELSE
    _REAL_TO_DWORD := DWORD#0;
  END_IF;
END_FUNCTION

FUNCTION _DWORD_TO_REAL:REAL
	VAR_INPUT
		IN :	DWORD;
	END_VAR

	_DWORD_TO_REAL := UDINT_TO_REAL(DWORD_TO_UDINT(IN));

END_FUNCTION

FUNCTION MULTIME:TIME
	VAR_INPUT
		T :	TIME;
		M :	REAL;
	END_VAR

	multime := DWORD_TO_TIME(_REAL_TO_DWORD(_DWORD_TO_REAL(TIME_TO_DWORD(t))*M));
END_FUNCTION

PROGRAM program0
  VAR
    LocalVar0 : TIME;
	LocalVar1 : REAL;
	LocalOUT  : TIME;
  END_VAR
  	LocalOUT := MULTIME(LocalVar0, LocalVar1);
END_PROGRAM

CONFIGURATION Config0
  RESOURCE Res0 ON PLC
    TASK task0(INTERVAL := T#20ms,PRIORITY := 0);
    PROGRAM instance0 WITH task0 : program0;
  END_RESOURCE
END_CONFIGURATION

(* ---- MUX_2.ST ---- *)
FUNCTION MUX_2:BOOL

	VAR_INPUT
		D0 :	BOOL;
		D1 :	BOOL;
		A0 :	BOOL;
	END_VAR

	MUX_2 := SEL(A0, D0, D1);

END_FUNCTION

PROGRAM program0
	VAR
		D0 :	BOOL;
		D1 :	BOOL;
		A0 :	BOOL;
		OUT : BOOL;
	END_VAR

	OUT := MUX_2(D0, D1, A0);

END_PROGRAM

CONFIGURATION Config0

	RESOURCE Res0 ON PLC
		TASK task0(INTERVAL := T#20ms,PRIORITY := 0);
		PROGRAM instance0 WITH task0 : program0;
	END_RESOURCE

END_CONFIGURATION

(* ---- MUX_4.ST ---- *)
FUNCTION MUX_4:BOOL

	VAR_INPUT
		D0 :	BOOL;
		D1 :	BOOL;
		D2 :	BOOL;
		D3 :	BOOL;
		A0 :	BOOL;
		A1 :	BOOL;
	END_VAR

	IF A1 THEN
		MUX_4 := SEL(A0, D2, D3);
	ELSE
		MUX_4 := SEL(A0, D0, D1);
	END_IF;

END_FUNCTION

PROGRAM program0
	VAR
		D0 :	BOOL;
		D1 :	BOOL;
		D2 :	BOOL;
		D3 :	BOOL;
		A0 :	BOOL;
		A1 :	BOOL;

		OUT : BOOL;
	END_VAR

	OUT := MUX_4(D0, D1, D2, D3, A0, A1);

END_PROGRAM

CONFIGURATION Config0

	RESOURCE Res0 ON PLC
		TASK task0(INTERVAL := T#20ms,PRIORITY := 0);
		PROGRAM instance0 WITH task0 : program0;
	END_RESOURCE

END_CONFIGURATION

(* ---- MUX_R2.ST ---- *)
FUNCTION MUX_R2:REAL

	VAR_INPUT
		IN0 :	REAL;
		IN1 :	REAL;
		A :	BOOL;
	END_VAR

	MUX_R2 := SEL(A, IN0, IN1);

END_FUNCTION

PROGRAM program0
	VAR
		IN0 :	REAL;
		IN1 :	REAL;
		A :	BOOL;

		OUT : REAL;
	END_VAR

	OUT := MUX_R2(IN0, IN1, A);

END_PROGRAM

CONFIGURATION Config0

	RESOURCE Res0 ON PLC
		TASK task0(INTERVAL := T#20ms,PRIORITY := 0);
		PROGRAM instance0 WITH task0 : program0;
	END_RESOURCE

END_CONFIGURATION

(* ---- MUX_R4.ST ---- *)
FUNCTION MUX_R4:REAL

	VAR_INPUT
		IN0 :	REAL;
		IN1 :	REAL;
		IN2 :	REAL;
		IN3 :	REAL;
		A0 :	BOOL;
		A1 :	BOOL;
	END_VAR

	IF A1 THEN
		MUX_R4 := SEL(A0, IN2, IN3);
	ELSE
		MUX_R4 := SEL(A0, IN0, IN1);
	END_IF;

END_FUNCTION

PROGRAM program0
	VAR
		IN0 :	REAL;
		IN1 :	REAL;
		IN2 :	REAL;
		IN3 :	REAL;
		A0 :	BOOL;
		A1 :	BOOL;

		OUT : REAL;
	END_VAR

	OUT := MUX_R4(IN0, IN1, IN2, IN3, A0, A1);

END_PROGRAM

CONFIGURATION Config0

	RESOURCE Res0 ON PLC
		TASK task0(INTERVAL := T#20ms,PRIORITY := 0);
		PROGRAM instance0 WITH task0 : program0;
	END_RESOURCE

END_CONFIGURATION

(* ---- NEGX.ST ---- *)
FUNCTION NEGX:REAL

	VAR_INPUT
		X :	REAL;
	END_VAR

	NEGX := -X;

END_FUNCTION

PROGRAM program0
	VAR
		_X : REAL;
		OUT : REAL;
	END_VAR

	OUT := NEGX(_X);
END_PROGRAM

CONFIGURATION Config0

	RESOURCE Res0 ON PLC
		TASK task0(INTERVAL := T#20ms,PRIORITY := 0);
		PROGRAM instance0 WITH task0 : program0;
	END_RESOURCE

END_CONFIGURATION

(* ---- NETWORK_VERSION.ST ---- *)
FUNCTION _INT_TO_UDINT:UDINT
	VAR_INPUT
		IN :	INT;
	END_VAR

	_INT_TO_UDINT := DINT_TO_UDINT(INT_TO_DINT(IN));
END_FUNCTION

FUNCTION SET_DATE:UDINT

	VAR_INPUT
		YEAR :	INT;
		MONTH :	INT;
		DAY :	INT;
	END_VAR

	VAR
		count :	INT;
	END_VAR

	IF month > 2 THEN
		count := (month - 1) * 30;
		IF month > 7 THEN
			count := count + DWORD_TO_INT(SHR(DINT_TO_DWORD(INT_TO_DINT(month) - INT_TO_DINT(3)),1));
		ELSE
			count := count + DWORD_TO_INT(SHR(DINT_TO_DWORD(INT_TO_DINT(month) - INT_TO_DINT(4)),1));
		END_IF;
		IF SHL(INT_TO_WORD(year),14) = WORD#0 THEN
			count := count + 1;
		END_IF;
	ELSE
		count := (month - 1) * 31;
	END_IF;
	SET_DATE := (_INT_TO_UDINT(count + day - 1) + DWORD_TO_UDINT(SHR(UDINT_TO_DWORD(_INT_TO_UDINT(year) * UDINT#1461 - UDINT#2878169), 2))) * UDINT#86400;

END_FUNCTION

FUNCTION NETWORK_VERSION:DWORD

	VAR_INPUT
		IN :	BOOL;
	END_VAR

	IF in THEN
		NETWORK_VERSION := UDINT_TO_DWORD(set_Date(2011,12,01));
	ELSE
		NETWORK_VERSION := DWORD#121;
	END_IF;

END_FUNCTION

PROGRAM program0
	VAR
		IN :	BOOL;
		CEIL5_OUT : DWORD;
	END_VAR

  	CEIL5_OUT := NETWORK_VERSION(IN);
END_PROGRAM

CONFIGURATION Config0

  RESOURCE Res0 ON PLC
    TASK task0(INTERVAL := T#20ms,PRIORITY := 0);
    PROGRAM instance0 WITH task0 : program0;
  END_RESOURCE
END_CONFIGURATION

(* ---- OFFSET.ST ---- *)
FUNCTION _OFFSET:REAL

	VAR_INPUT
		X :	REAL;
		O1 :	BOOL;
		O2 :	BOOL;
		O3 :	BOOL;
		O4 :	BOOL;
		D :	BOOL;
		OFFSET_1 :	REAL;
		OFFSET_2 :	REAL;
		OFFSET_3 :	REAL;
		OFFSET_4 :	REAL;
		DEFAULT :	REAL;
	END_VAR

	IF D THEN _Offset := default; ELSE _Offset := X; END_IF;
	IF O1 THEN _Offset := _Offset + offset_1; END_IF;
	IF O2 THEN _Offset := _Offset + offset_2; END_IF;
	IF O3 THEN _Offset := _Offset + offset_3; END_IF;
	IF O4 THEN _Offset := _Offset + offset_4; END_IF;

END_FUNCTION

PROGRAM program0

	VAR
		X :	REAL;
		O1 :	BOOL;
		O2 :	BOOL;
		O3 :	BOOL;
		O4 :	BOOL;
		D :	BOOL;
		OFFSET_1 :	REAL;
		OFFSET_2 :	REAL;
		OFFSET_3 :	REAL;
		OFFSET_4 :	REAL;
		DEFAULT :	REAL;
		OUT : REAL;
	END_VAR

	OUT := _OFFSET(X, O1, O2, O3, O4, D, OFFSET_1, OFFSET_2, OFFSET_3, OFFSET_4, DEFAULT);
END_PROGRAM

CONFIGURATION Config0

	RESOURCE Res0 ON PLC
		TASK task0(INTERVAL := T#20ms,PRIORITY := 0);
		PROGRAM instance0 WITH task0 : program0;
	END_RESOURCE

END_CONFIGURATION

(* ---- OFFSET2.ST ---- *)
FUNCTION OFFSET2:REAL

	VAR_INPUT
		X :	REAL;
		O1 :	BOOL;
		O2 :	BOOL;
		O3 :	BOOL;
		O4 :	BOOL;
		D :	BOOL;
		OFFSET_1 :	REAL;
		OFFSET_2 :	REAL;
		OFFSET_3 :	REAL;
		OFFSET_4 :	REAL;
		DEFAULT :	REAL;
	END_VAR

	IF D THEN Offset2 := default; ELSE Offset2 := X; END_IF;
	IF O4 THEN Offset2 := Offset2 + offset_4;
	ELSIF O3 THEN Offset2 := Offset2 + offset_3;
	ELSIF O2 THEN Offset2 := Offset2 + offset_2;
	ELSIF O1 THEN Offset2 := Offset2 + offset_1;
	END_IF;

END_FUNCTION

PROGRAM program0
	VAR
		X :	REAL;
		O1 :	BOOL;
		O2 :	BOOL;
		O3 :	BOOL;
		O4 :	BOOL;
		D :	BOOL;
		OFFSET_1 :	REAL;
		OFFSET_2 :	REAL;
		OFFSET_3 :	REAL;
		OFFSET_4 :	REAL;
		DEFAULT :	REAL;
		OUT : REAL;
	END_VAR

	OUT := OFFSET2(X, O1, O2, O3, O4, D, OFFSET_1, OFFSET_2, OFFSET_3, OFFSET_4, DEFAULT);
END_PROGRAM

CONFIGURATION Config0

	RESOURCE Res0 ON PLC
		TASK task0(INTERVAL := T#20ms,PRIORITY := 0);
		PROGRAM instance0 WITH task0 : program0;
	END_RESOURCE

END_CONFIGURATION

(* ---- OM_TO_F.ST ---- *)
FUNCTION OM_TO_F:REAL

	VAR_INPUT
		OM :	REAL;
	END_VAR

	OM_to_F := OM / 6.283185307179586476;

END_FUNCTION

PROGRAM program0
	VAR
		OM : REAL;
		OUT : REAL;
	END_VAR

	OUT := OM_TO_F(OM);
END_PROGRAM

CONFIGURATION Config0

	RESOURCE Res0 ON PLC
		TASK task0(INTERVAL := T#20ms,PRIORITY := 0);
		PROGRAM instance0 WITH task0 : program0;
	END_RESOURCE

END_CONFIGURATION

(* ---- OSCAT_VERSION.ST ---- *)
FUNCTION _INT_TO_UDINT:UDINT
	VAR_INPUT
		IN :	INT;
	END_VAR

	_INT_TO_UDINT := DINT_TO_UDINT(INT_TO_DINT(IN));
END_FUNCTION

FUNCTION SET_DATE:UDINT

	VAR_INPUT
		YEAR :	INT;
		MONTH :	INT;
		DAY :	INT;
	END_VAR

	VAR
		count :	INT;
	END_VAR

	IF month > 2 THEN
		count := (month - 1) * 30;
		IF month > 7 THEN
			count := count + DWORD_TO_INT(SHR(DINT_TO_DWORD(INT_TO_DINT(month) - INT_TO_DINT(3)),1));
		ELSE
			count := count + DWORD_TO_INT(SHR(DINT_TO_DWORD(INT_TO_DINT(month) - INT_TO_DINT(4)),1));
		END_IF;
		IF SHL(INT_TO_WORD(year),14) = WORD#0 THEN
			count := count + 1;
		END_IF;
	ELSE
		count := (month - 1) * 31;
	END_IF;
	SET_DATE := (_INT_TO_UDINT(count + day - 1) + DWORD_TO_UDINT(SHR(UDINT_TO_DWORD(_INT_TO_UDINT(year) * UDINT#1461 - UDINT#2878169), 2))) * UDINT#86400;

END_FUNCTION

FUNCTION OSCAT_VERSION:DWORD

	VAR_INPUT
		IN :	BOOL;
	END_VAR

	IF in THEN
		Oscat_version := UDINT_TO_DWORD(set_Date(2012,01,02));
	ELSE
		Oscat_version := DWORD#333;
	END_IF;

END_FUNCTION

PROGRAM program0
	VAR
		IN :	BOOL;
		OUT : DWORD;
	END_VAR

	OUT := OSCAT_VERSION(IN);
END_PROGRAM

CONFIGURATION Config0

	RESOURCE Res0 ON PLC
		TASK task0(INTERVAL := T#20ms,PRIORITY := 0);
		PROGRAM instance0 WITH task0 : program0;
	END_RESOURCE

END_CONFIGURATION

(* ---- PARITY.ST ---- *)
FUNCTION BIT_OF_DWORD : BOOL

	VAR_INPUT
		IN : DWORD;
		N : INT;
	END_VAR

	BIT_OF_DWORD := (SHR(in,N) AND 16#00000001) > 0;

END_FUNCTION

FUNCTION PARITY:BOOL

	VAR_INPUT
		IN :	DWORD;
	END_VAR

	VAR
		in2 :	DWORD;
	END_VAR

	in2:=in;
	WHILE in2 > DWORD#0 DO
		parity := parity XOR BIT_OF_DWORD(in2,0) XOR BIT_OF_DWORD(in2,1) XOR BIT_OF_DWORD(in2,2) XOR BIT_OF_DWORD(in2,3);
		in2 := SHR(in2,4);
	END_WHILE;

END_FUNCTION

PROGRAM program0
	VAR
		IN : DWORD;
		OUT : BOOL;
	END_VAR

	OUT := PARITY(IN);
END_PROGRAM

CONFIGURATION Config0

	RESOURCE Res0 ON PLC
		TASK task0(INTERVAL := T#20ms,PRIORITY := 0);
		PROGRAM instance0 WITH task0 : program0;
	END_RESOURCE

END_CONFIGURATION

(* ---- PERIOD.ST ---- *)
FUNCTION LEAP_OF_DATE:BOOL

	VAR_INPUT
		IDATE :	UDINT;
	END_VAR

	LEAP_OF_DATE := SHL(UDINT_TO_DWORD((idate + UDINT#43200) / UDINT#31557600), 30) = DWORD#16#80000000;
END_FUNCTION

FUNCTION DAY_OF_YEAR:INT
	VAR_INPUT
		IDATE :	UDINT;
	END_VAR

	DAY_OF_YEAR := UDINT_TO_INT(((idate) / UDINT#86400) MOD UDINT#1461);
	IF DAY_OF_YEAR > 729 THEN
		IF DAY_OF_YEAR > 1095 THEN DAY_OF_YEAR := DAY_OF_YEAR - 1095; ELSE DAY_OF_YEAR := DAY_OF_YEAR - 729; END_IF;
	ELSIF DAY_OF_YEAR > 364 THEN
		DAY_OF_YEAR := DAY_OF_YEAR - 364;
	ELSE
		DAY_OF_YEAR := DAY_OF_YEAR + 1;
	END_IF;
END_FUNCTION

FUNCTION PERIOD:BOOL

	VAR
		day1 :	INT;
		day2 :	INT;
		dayx :	INT;
	END_VAR

	VAR_INPUT
		D1 :	UDINT;
		Dx :	UDINT;
		D2 :	UDINT;
	END_VAR

	day1 := day_of_year(d1);
	day2 := day_of_year(d2);
	dayx := day_of_year(dx);
	IF NOT leap_of_Date(dx) AND dayx > 58 THEN dayx := dayx + 1; END_IF;
	IF NOT leap_of_Date(d1) AND day1 > 58 THEN day1 := day1 + 1; END_IF;
	IF NOT leap_of_Date(d2) AND day2 > 58 THEN day2 := day2 + 1; END_IF;

	IF day2 < day1 THEN
		(* the period spans over the new year *)
		period := dayx <= day2 OR dayx >= day1;
	ELSE
		period := dayx >= day1 AND dayx <= day2;
	END_IF;

END_FUNCTION

PROGRAM program0
	VAR
		D1 :	UDINT;
		Dx :	UDINT;
		D2 :	UDINT;

		OUT : BOOL;
	END_VAR

	OUT := PERIOD(D1, Dx, D2);
END_PROGRAM

CONFIGURATION Config0

	RESOURCE Res0 ON PLC
		TASK task0(INTERVAL := T#20ms,PRIORITY := 0);
		PROGRAM instance0 WITH task0 : program0;
	END_RESOURCE

END_CONFIGURATION

(* ---- PT_TO_F.ST ---- *)
FUNCTION _DWORD_TO_REAL:REAL
	VAR_INPUT
		IN :	DWORD;
	END_VAR

	_DWORD_TO_REAL := UDINT_TO_REAL(DWORD_TO_UDINT(IN));

END_FUNCTION

FUNCTION PT_TO_F:REAL

	VAR_INPUT
		PT :	TIME;
	END_VAR

	PT_TO_F := 1000.0 / _DWORD_TO_REAL(TIME_TO_DWORD(PT));

END_FUNCTION

PROGRAM program0
  VAR
    PT : TIME;
    OUT : REAL;
  END_VAR

  OUT := PT_TO_F(PT);
END_PROGRAM

CONFIGURATION Config0

  RESOURCE Res0 ON PLC
    TASK task0(INTERVAL := T#20ms,PRIORITY := 0);
    PROGRAM instance0 WITH task0 : program0;
  END_RESOURCE
END_CONFIGURATION

(* ---- RAD.ST ---- *)
FUNCTION FLOOR2 : DINT
	VAR_INPUT
		x : REAL;
	END_VAR

	FLOOR2 := REAL_TO_DINT(X);
	IF DINT_TO_REAL(FLOOR2) > X THEN
		FLOOR2 := FLOOR2 - DINT#1;
	END_IF;

END_FUNCTION

FUNCTION MODR: REAL

	VAR_INPUT
		IN :	REAL;
		DIVI :	REAL;
	END_VAR

	IF divi = 0.0 THEN
		MODR := 0.0;
	ELSE
		MODR := in - DINT_TO_REAL(FLOOR2(in / divi)) * divi;
	END_IF;

END_FUNCTION

FUNCTION RAD:REAL

	VAR_INPUT
		DEG :	REAL;
	END_VAR

	RAD := MODR(0.0174532925199433 * DEG , 6.283185307179586476);

END_FUNCTION

PROGRAM program0

	VAR
		DEG :	REAL;
		CEIL5_OUT : REAL;
	END_VAR

	CEIL5_OUT := RAD(DEG);

END_PROGRAM

CONFIGURATION Config0

	RESOURCE Res0 ON PLC
		TASK task0(INTERVAL := T#20ms,PRIORITY := 0);
		PROGRAM instance0 WITH task0 : program0;
	END_RESOURCE

END_CONFIGURATION

(* ---- RANGE_TO_BYTE.ST ---- *)
FUNCTION TRUNC_REAL:REAL

	VAR_INPUT
		IN :	REAL;
	END_VAR

	TRUNC_REAL := UDINT_TO_REAL(DINT_TO_UDINT(TRUNC(IN)));
END_FUNCTION

FUNCTION RANGE_TO_BYTE:BYTE

	VAR_INPUT
		X :	REAL;
		LOW :	REAL;
		HIGH :	REAL;
	END_VAR

	Range_to_Byte := REAL_TO_BYTE(TRUNC_REAL((LIMIT(low,X,high)-low) * 255.0 / (high - low)));

END_FUNCTION

PROGRAM program0

	VAR
		X :	REAL;
		LOW :	REAL;
		HIGH :	REAL;

        OUT :	BYTE;
	END_VAR
	OUT := RANGE_TO_BYTE(X, LOW, HIGH);

END_PROGRAM

CONFIGURATION Config0

	RESOURCE Res0 ON PLC
		TASK task0(INTERVAL := T#20ms,PRIORITY := 0);
		PROGRAM instance0 WITH task0 : program0;
	END_RESOURCE

END_CONFIGURATION

(* ---- RANGE_TO_WORD.ST ---- *)
FUNCTION TRUNC_REAL:REAL

	VAR_INPUT
		IN :	REAL;
	END_VAR

	TRUNC_REAL := UDINT_TO_REAL(DINT_TO_UDINT(TRUNC(IN)));
END_FUNCTION

FUNCTION RANGE_TO_WORD:WORD

	VAR_INPUT
		X :	REAL;
		LOW :	REAL;
		HIGH :	REAL;
	END_VAR

	Range_to_Word := REAL_TO_WORD(TRUNC_REAL((LIMIT(low,X,high)-low) * 65535.0 / (high - low)));

END_FUNCTION

PROGRAM program0

	VAR
		X :	REAL;
		LOW :	REAL;
		HIGH :	REAL;

        OUT :	WORD;
	END_VAR
	OUT := RANGE_TO_WORD(X, LOW, HIGH);

END_PROGRAM

CONFIGURATION Config0

	RESOURCE Res0 ON PLC
		TASK task0(INTERVAL := T#20ms,PRIORITY := 0);
		PROGRAM instance0 WITH task0 : program0;
	END_RESOURCE

END_CONFIGURATION

(* ---- REAL_TO_TIME.ST ---- *)
FUNCTION _REAL_TO_UDINT:UDINT
  VAR_INPUT
    X :	REAL;
  END_VAR

  IF REAL_TO_UDINT(0.5) = UDINT#1 THEN
    _REAL_TO_UDINT := REAL_TO_UDINT(x);
  ELSIF X > 0.0 THEN
    _REAL_TO_UDINT := REAL_TO_UDINT(x+0.5);
  ELSIF X < 0.0 THEN
    _REAL_TO_UDINT := REAL_TO_UDINT(x-0.5);
  ELSE
    _REAL_TO_UDINT := UDINT#0;
  END_IF;
END_FUNCTION

FUNCTION REAL_TO_TIME2:TIME
	VAR_INPUT
		IN :	REAL;
	END_VAR

	REAL_TO_TIME2 := DINT_TO_TIME(UDINT_TO_DINT(_REAL_TO_UDINT(IN)));
END_FUNCTION

PROGRAM program0
  VAR
    LocalVar0 : REAL;
    LocalOUT  : TIME;
  END_VAR

  LocalOUT := REAL_TO_TIME2(LocalVar0);
END_PROGRAM

CONFIGURATION Config0
  RESOURCE Res0 ON PLC
    TASK task0(INTERVAL := T#20ms,PRIORITY := 0);
    PROGRAM instance0 WITH task0 : program0;
  END_RESOURCE
END_CONFIGURATION

(* ---- REFLECT.ST ---- *)
FUNCTION REFLECT:DWORD
	VAR_INPUT
		D :	DWORD;
		L :	INT;
	END_VAR

	VAR
		i :	INT;
		_d :	DWORD;
	END_VAR

	REFLECT := DWORD#0;
	_d := D;
	FOR i := 1 TO L DO
		REFLECT := SHL(REFLECT, 1) OR BOOL_TO_DWORD((_d AND DWORD#2#0000_0001) > DWORD#0); (* D.0 *)
		_d := SHR(_d, 1);
	END_FOR;
	REFLECT := REFLECT OR SHL(_d, L);
END_FUNCTION

PROGRAM program0
  VAR
    LocalVar0 : DWORD;
	LocalVar1 : INT;
	LocalOUT  : DWORD;
  END_VAR
  	LocalOUT := REFLECT(LocalVar0, LocalVar1);
END_PROGRAM

CONFIGURATION Config0
  RESOURCE Res0 ON PLC
    TASK task0(INTERVAL := T#20ms,PRIORITY := 0);
    PROGRAM instance0 WITH task0 : program0;
  END_RESOURCE
END_CONFIGURATION

(* ---- REFRACTION.ST ---- *)
FUNCTION REFRACTION:REAL

	VAR_INPUT
		ELEV :	REAL;
	END_VAR

	VAR
		tmp :	REAL;
	END_VAR

	tmp := LIMIT(-1.9, elev, 80.0);
	REFRACTION := 0.0174532925199433 / TAN(0.0174532925199433 * (tmp + 10.3 / (tmp + 5.11)));

END_FUNCTION

PROGRAM program0

	VAR
		ELEV :	REAL;

		OUT :	REAL;
	END_VAR
	OUT := REFRACTION(ELEV);

END_PROGRAM

CONFIGURATION Config0

	RESOURCE Res0 ON PLC
		TASK task0(INTERVAL := T#20ms,PRIORITY := 0);
		PROGRAM instance0 WITH task0 : program0;
	END_RESOURCE

END_CONFIGURATION

(* ---- RES_NI.ST ---- *)
FUNCTION RES_NI:REAL

	VAR_INPUT
		T :	REAL;
		R0 :	REAL;
	END_VAR

	VAR
		T2 :	REAL;
	END_VAR

	T2 := T*T;
	Res_NI := R0 + 0.5485*T + 0.665E-3*T2 + 2.805E-9*T2*T2;

END_FUNCTION

PROGRAM program0

	VAR
		T :	REAL;
		R0 :	REAL;

		OUT :	REAL;
	END_VAR
	OUT := RES_NI(T, R0);

END_PROGRAM

CONFIGURATION Config0

	RESOURCE Res0 ON PLC
		TASK task0(INTERVAL := T#20ms,PRIORITY := 0);
		PROGRAM instance0 WITH task0 : program0;
	END_RESOURCE

END_CONFIGURATION

(* ---- RES_NTC.ST ---- *)
FUNCTION RES_NTC:REAL

	VAR_INPUT
		T :	REAL;
		RN :	REAL;
		B :	REAL;
	END_VAR

	RES_NTC := RN * EXP(B * (1.0 / (T+273.15) - 0.00335401643468053));

END_FUNCTION

PROGRAM program0

	VAR
		T :	REAL;
		RN :	REAL;
		B :	REAL;

		OUT :	REAL;
	END_VAR
		OUT := RES_NTC(T, RN, B);

END_PROGRAM

CONFIGURATION Config0

	RESOURCE Res0 ON PLC
		TASK task0(INTERVAL := T#20ms,PRIORITY := 0);
		PROGRAM instance0 WITH task0 : program0;
	END_RESOURCE

END_CONFIGURATION

(* ---- RES_PT.ST ---- *)
FUNCTION RES_PT:REAL
	VAR_INPUT
		T :	REAL;
		R0 :	REAL;
	END_VAR

	VAR
		T2 :	REAL;
	END_VAR

	T2 := T * T;

	IF T >= 0.0 THEN
		RES_PT := R0 * ( 1.0 + 3.90802E-3 * T + -5.802E-7 * T2);
	ELSE
		RES_PT := R0 * ( 1.0 + 3.90802E-3 * T + -5.802E-7 * T2 + -4.27350E-12 * (T - 100.0) * T2 * T);
	END_IF;

END_FUNCTION

PROGRAM program0
  	VAR
		T :	REAL;
		R0 : REAL;
		CEIL5_OUT : REAL;
  	END_VAR

  	CEIL5_OUT := RES_PT(T, R0);
END_PROGRAM

CONFIGURATION Config0
	RESOURCE Res0 ON PLC
		TASK task0(INTERVAL := T#20ms,PRIORITY := 0);
		PROGRAM instance0 WITH task0 : program0;
	END_RESOURCE
END_CONFIGURATION

(* ---- RES_SI.ST ---- *)
FUNCTION RES_SI:REAL

	VAR_INPUT
		T :	REAL;
		_RS :	REAL;
		TS :	REAL;
	END_VAR

	VAR
		TX :	REAL;
	END_VAR

	TX := T - TS;
	RES_SI := _RS * ( 1.0 + 7.64E-3 * TX + 1.66E-5 * TX * TX);

END_FUNCTION

PROGRAM program0

	VAR
		T :	REAL;
		_RS :	REAL;
		TS :	REAL;

		OUT :	REAL;
	END_VAR
		OUT := RES_SI(T, _RS, TS);

END_PROGRAM

CONFIGURATION Config0

	RESOURCE Res0 ON PLC
		TASK task0(INTERVAL := T#20ms,PRIORITY := 0);
		PROGRAM instance0 WITH task0 : program0;
	END_RESOURCE

END_CONFIGURATION

(* ---- REVERSE.ST ---- *)
FUNCTION REVERSE:BYTE
VAR_INPUT
	IN :	BYTE;
END_VAR

reverse := SHL(in,7) OR SHR(in,7) OR (ROR(in,3) AND BYTE#2#01000100) OR (ROL(in,3) AND BYTE#2#00100010)
	OR (SHL(in,1) AND BYTE#2#00010000) OR (SHR(in,1) AND BYTE#2#00001000);

END_FUNCTION

PROGRAM program0
  VAR
    LocalVar0 : BYTE;
	LocalOUT  : BYTE;
  END_VAR
  	LocalOUT := REVERSE(LocalVar0);
END_PROGRAM

CONFIGURATION Config0
  RESOURCE Res0 ON PLC
    TASK task0(INTERVAL := T#20ms,PRIORITY := 0);
    PROGRAM instance0 WITH task0 : program0;
  END_RESOURCE
END_CONFIGURATION

(* ---- RND.ST ---- *)
FUNCTION CEIL:INT

	VAR_INPUT
		X :	REAL;
	END_VAR

	CEIL := REAL_TO_INT(x);
	IF INT_TO_REAL(CEIL) < X THEN
			CEIL := CEIL + 1;
	END_IF;

END_FUNCTION

FUNCTION BIT_OF_DWORD : BOOL

	VAR_INPUT
		IN : DWORD;
		N : INT;
	END_VAR

	BIT_OF_DWORD := (SHR(in,N) AND 16#00000001) > 0;

END_FUNCTION

FUNCTION EXPN:REAL

	VAR_INPUT
		X :	REAL;
		N :	INT;
	END_VAR

	VAR
		N_word :	WORD;
		X_tmp :	REAL;
		sign :	BOOL;
	END_VAR

	N_word := INT_TO_WORD(N);
	X_tmp := X;
	sign := BIT_OF_DWORD(WORD_TO_DWORD(N_word),15);
	N_word := INT_TO_WORD(ABS(N));
	IF BIT_OF_DWORD(WORD_TO_DWORD(N_word),0) THEN expn := X_tmp; ELSE expn := 1.0; END_IF;    (* N_word.X0 *)
	N_word := SHR(N_word,1);
	WHILE N_word > WORD#0 DO
		X_tmp := X_tmp * X_tmp;
		IF BIT_OF_DWORD(WORD_TO_DWORD(N_word),0) THEN expn := expn * X_tmp; END_IF;       (* N_word.X0 *)
		N_word := SHR(N_word,1);
	END_WHILE;
	IF sign THEN EXPN := 1.0 / EXPN; END_IF;

END_FUNCTION

FUNCTION _REAL_TO_DINT:DINT
	VAR_INPUT
		X :	REAL;
	END_VAR

	IF REAL_TO_DINT(0.5) = DINT#1 THEN
		_REAL_TO_DINT := REAL_TO_DINT(x);
		RETURN;
	END_IF;

	IF X > 0.0 THEN
		_REAL_TO_DINT := REAL_TO_DINT(x+0.5);
	ELSIF X < 0.0 THEN
		_REAL_TO_DINT := REAL_TO_DINT(x-0.5);
	ELSE
		_REAL_TO_DINT := DINT#0;
	END_IF;
END_FUNCTION

FUNCTION RND:REAL

	VAR_INPUT
		X :	REAL;
		N :	INT;
	END_VAR

	VAR
		M :	REAL;
	END_VAR

	IF X = 0.0 THEN
		RND := 0.0;
	ELSE
		M := EXPN(10.0,N - CEIL(LOG(ABS(X))));
		RND := DINT_TO_REAL(_REAL_TO_DINT(X * M)) / M;
	END_IF;

END_FUNCTION

PROGRAM program0
	VAR
		IN : REAL;
		N :	INT;
		X :	REAL;
	END_VAR
		X := RND(IN, N);
END_PROGRAM

CONFIGURATION Config0

	RESOURCE Res0 ON PLC
		TASK task0(INTERVAL := T#20ms,PRIORITY := 0);
		PROGRAM instance0 WITH task0 : program0;
	END_RESOURCE

END_CONFIGURATION

(* ---- ROUND.ST ---- *)
FUNCTION _REAL_TO_DINT:DINT
	VAR_INPUT
		X :	REAL;
	END_VAR

	IF REAL_TO_DINT(0.5) = DINT#1 THEN
		_REAL_TO_DINT := REAL_TO_DINT(x);
		RETURN;
	END_IF;

	IF X > 0.0 THEN
		_REAL_TO_DINT := REAL_TO_DINT(x+0.5);
	ELSIF X < 0.0 THEN
		_REAL_TO_DINT := REAL_TO_DINT(x-0.5);
	ELSE
		_REAL_TO_DINT := DINT#0;
	END_IF;
END_FUNCTION

FUNCTION ROUND:REAL

	VAR_INPUT
		IN :	REAL;
		N :	INT;
	END_VAR

	VAR
		X :	REAL;
	END_VAR

	IF N < 4 THEN
		IF N < 2 THEN
			IF N = 0 THEN X := 1.0; ELSE X := 10.0; END_IF;
		ELSE
			IF N = 2 THEN X := 100.0; ELSE X := 1000.0; END_IF;
		END_IF;
	ELSE
		IF N < 6 THEN
			IF N = 4 THEN X := 10000.0; ELSE X := 100000.0; END_IF;
		ELSE
			IF N = 6 THEN X := 1000000.0; ELSE X := 10000000.0; END_IF;
		END_IF;
	END_IF;

	ROUND := DINT_TO_REAL(_REAL_TO_DINT(in * X)) / X;

END_FUNCTION

PROGRAM program0
	VAR
		IN : REAL;
		N :	INT;
		X :	REAL;
	END_VAR
		X := ROUND(IN, N);
END_PROGRAM

CONFIGURATION Config0

	RESOURCE Res0 ON PLC
		TASK task0(INTERVAL := T#20ms,PRIORITY := 0);
		PROGRAM instance0 WITH task0 : program0;
	END_RESOURCE

END_CONFIGURATION

(* ---- SCALE.ST ---- *)
FUNCTION SCALE:REAL

	VAR_INPUT
		X :	REAL;
		K :	REAL;
		O :	REAL;
		MX :	REAL;
		MN :	REAL;
	END_VAR

	SCALE := LIMIT(MN, X * K + O, MX);

END_FUNCTION

PROGRAM program0
  VAR
    X :	REAL;
	K :	REAL;
	O :	REAL;
	MX :	REAL;
	MN :	REAL;
    CEIL5_OUT : REAL;
  END_VAR

  CEIL5_OUT := SCALE(X, K, O, MX, MN);
END_PROGRAM

CONFIGURATION Config0

  RESOURCE Res0 ON PLC
    TASK task0(INTERVAL := T#20ms,PRIORITY := 0);
    PROGRAM instance0 WITH task0 : program0;
  END_RESOURCE
END_CONFIGURATION

(* ---- SCALE_B.ST ---- *)
FUNCTION _BYTE_TO_REAL:REAL
	VAR_INPUT
		IN :	BYTE;
	END_VAR

	_BYTE_TO_REAL := USINT_TO_REAL(BYTE_TO_USINT(IN));
END_FUNCTION

FUNCTION SCALE_B:REAL

	VAR_INPUT
		X :	BYTE;
		I_LO :	BYTE;
		I_HI :	BYTE;
		O_LO :	REAL;
		O_HI :	REAL;
	END_VAR

	IF I_HI = I_LO THEN
		SCALE_B := O_LO;
	ELSE
		SCALE_B := (O_HI - O_LO) / USINT_TO_REAL(BYTE_TO_USINT(I_HI) - BYTE_TO_USINT(I_LO)) * _BYTE_TO_REAL(LIMIT(I_LO,X,I_HI));
	END_IF;

END_FUNCTION

PROGRAM program0
  VAR
	X :	BYTE;
	I_LO :	BYTE;
	I_HI :	BYTE;
	O_LO :	REAL;
	O_HI :	REAL;
	CEIL5_OUT : REAL;
  END_VAR

  CEIL5_OUT := SCALE_B(X, I_LO, I_HI, O_LO, O_HI);

END_PROGRAM

CONFIGURATION Config0

  RESOURCE Res0 ON PLC
    TASK task0(INTERVAL := T#20ms,PRIORITY := 0);
    PROGRAM instance0 WITH task0 : program0;
  END_RESOURCE
END_CONFIGURATION

(* ---- SCALE_B2.ST ---- *)
FUNCTION _BYTE_TO_REAL:REAL
	VAR_INPUT
		IN :	BYTE;
	END_VAR

	_BYTE_TO_REAL := USINT_TO_REAL(BYTE_TO_USINT(IN));
END_FUNCTION

FUNCTION SCALE_B2:REAL
	VAR_INPUT
		IN1 :	BYTE;
		IN2 :	BYTE;
		K :	REAL;
		O :	REAL;
		IN1_MIN :	REAL;
		IN1_MAX :	REAL;
		IN2_MIN :	REAL;
		IN2_MAX :	REAL;
	END_VAR

	SCALE_B2 := 	(((in1_max - in1_min)* _BYTE_TO_REAL(in1) + (in2_max - in2_min)* _BYTE_TO_REAL(in2)) * 0.003921569 + in1_min + in2_min) * K + O;

END_FUNCTION

PROGRAM program0
  VAR
	IN1 :	BYTE;
	IN2 :	BYTE;
	K :	REAL;
	O :	REAL;
	IN1_MIN :	REAL;
	IN1_MAX :	REAL;
	IN2_MIN :	REAL;
	IN2_MAX :	REAL;
	CEIL5_OUT : REAL;
  END_VAR

  CEIL5_OUT := SCALE_B2(IN1, IN2, K, O, IN1_MIN, IN1_MAX, IN2_MIN, IN2_MAX);

END_PROGRAM

CONFIGURATION Config0

  RESOURCE Res0 ON PLC
    TASK task0(INTERVAL := T#20ms,PRIORITY := 0);
    PROGRAM instance0 WITH task0 : program0;
  END_RESOURCE
END_CONFIGURATION

(* ---- SCALE_B4.ST ---- *)
FUNCTION _BYTE_TO_REAL:REAL
	VAR_INPUT
		IN :	BYTE;
	END_VAR

	_BYTE_TO_REAL := USINT_TO_REAL(BYTE_TO_USINT(IN));
END_FUNCTION

FUNCTION SCALE_B4:REAL

	VAR_INPUT
		IN1 :	BYTE;
		IN2 :	BYTE;
		IN3 :	BYTE;
		IN4 :	BYTE;
		K :	REAL;
		O :	REAL;
		IN1_MIN :	REAL;
		IN1_MAX :	REAL;
		IN2_MIN :	REAL;
		IN2_MAX :	REAL;
		IN3_MIN :	REAL;
		IN3_MAX :	REAL;
		IN4_MIN :	REAL;
		IN4_MAX :	REAL;
	END_VAR

	SCALE_B4 := 	(((in1_max - in1_min)* _BYTE_TO_REAL(in1) + (in2_max - in2_min)* _BYTE_TO_REAL(in2) + (in3_max - in3_min)* _BYTE_TO_REAL(in3) + (in4_max - in4_min)* _BYTE_TO_REAL(in4))* 0.003921569 + in1_min + in2_min + in3_min + in4_min) * K + O;

END_FUNCTION

PROGRAM program0
  VAR
	IN1 :	BYTE;
	IN2 :	BYTE;
	IN3 :	BYTE;
	IN4 :	BYTE;
	K :	REAL;
	O :	REAL;
	IN1_MIN :	REAL;
	IN1_MAX :	REAL;
	IN2_MIN :	REAL;
	IN2_MAX :	REAL;
	IN3_MIN :	REAL;
	IN3_MAX :	REAL;
	IN4_MIN :	REAL;
	IN4_MAX :	REAL;
	CEIL5_OUT : REAL;
  END_VAR

  CEIL5_OUT := SCALE_B4(IN1, IN2, IN3, IN4, K, O, IN1_MIN, IN1_MAX, IN2_MIN, IN2_MAX, IN3_MIN, IN3_MAX, IN4_MIN, IN4_MAX);

END_PROGRAM

CONFIGURATION Config0

  RESOURCE Res0 ON PLC
    TASK task0(INTERVAL := T#20ms,PRIORITY := 0);
    PROGRAM instance0 WITH task0 : program0;
  END_RESOURCE
END_CONFIGURATION

(* ---- SCALE_B8.ST ---- *)
FUNCTION _BYTE_TO_REAL:REAL
	VAR_INPUT
		IN :	BYTE;
	END_VAR

	_BYTE_TO_REAL := USINT_TO_REAL(BYTE_TO_USINT(IN));
END_FUNCTION

FUNCTION SCALE_B8:REAL
	VAR_INPUT
		IN1 :	BYTE;
		IN2 :	BYTE;
		IN3 :	BYTE;
		IN4 :	BYTE;
		IN5 :	BYTE;
		IN6 :	BYTE;
		IN7 :	BYTE;
		IN8 :	BYTE;
		K :	REAL;
		O :	REAL;
		IN1_MIN :	REAL;
		IN1_MAX :	REAL;
		IN2_MIN :	REAL;
		IN2_MAX :	REAL;
		IN3_MIN :	REAL;
		IN3_MAX :	REAL;
		IN4_MIN :	REAL;
		IN4_MAX :	REAL;
		IN5_MIN :	REAL;
		IN5_MAX :	REAL;
		IN6_MIN :	REAL;
		IN6_MAX :	REAL;
		IN7_MIN :	REAL;
		IN7_MAX :	REAL;
		IN8_MIN :	REAL;
		IN8_MAX :	REAL;
	END_VAR

	SCALE_B8 := 	(((in1_max - in1_min)* _BYTE_TO_REAL(in1) + (in2_max - in2_min)* _BYTE_TO_REAL(in2) + (in3_max - in3_min)* _BYTE_TO_REAL(in3) + (in4_max - in4_min)* _BYTE_TO_REAL(in4) +
					(in5_max - in5_min)* _BYTE_TO_REAL(in5) + (in6_max - in6_min)* _BYTE_TO_REAL(in6) + (in7_max - in7_min)* _BYTE_TO_REAL(in7) + (in8_max - in8_min)* _BYTE_TO_REAL(in8)) * 0.003921569
					+ in1_min + in2_min + in3_min + in4_min + in5_min + in6_min + in7_min + in8_min) * K + O;

END_FUNCTION

PROGRAM program0
  	VAR
		IN1 :	BYTE;
		IN2 :	BYTE;
		IN3 :	BYTE;
		IN4 :	BYTE;
		IN5 :	BYTE;
		IN6 :	BYTE;
		IN7 :	BYTE;
		IN8 :	BYTE;
		K :	REAL;
		O :	REAL;
		IN1_MIN :	REAL;
		IN1_MAX :	REAL;
		IN2_MIN :	REAL;
		IN2_MAX :	REAL;
		IN3_MIN :	REAL;
		IN3_MAX :	REAL;
		IN4_MIN :	REAL;
		IN4_MAX :	REAL;
		IN5_MIN :	REAL;
		IN5_MAX :	REAL;
		IN6_MIN :	REAL;
		IN6_MAX :	REAL;
		IN7_MIN :	REAL;
		IN7_MAX :	REAL;
		IN8_MIN :	REAL;
		IN8_MAX :	REAL;
		CEIL5_OUT : REAL;
  	END_VAR

  	CEIL5_OUT := SCALE_B8(IN1, IN2, IN3, IN4, IN5, IN6, IN7, IN8, K, O, IN1_MIN, IN1_MAX, IN2_MIN, IN2_MAX, IN3_MIN, IN3_MAX, IN4_MIN, IN4_MAX, IN5_MIN, IN5_MAX, IN6_MIN, IN6_MAX, IN7_MIN, IN7_MAX, IN8_MIN, IN8_MAX);

	END_PROGRAM

CONFIGURATION Config0

	RESOURCE Res0 ON PLC
		TASK task0(INTERVAL := T#20ms,PRIORITY := 0);
		PROGRAM instance0 WITH task0 : program0;
	END_RESOURCE

END_CONFIGURATION

(* ---- SCALE_D.ST ---- *)
FUNCTION SCALE_D:REAL
	VAR_INPUT
		X :	DWORD;
		I_LO :	DWORD;
		I_HI :	DWORD;
		O_LO :	REAL;
		O_HI :	REAL;
	END_VAR
	IF I_HI = I_LO THEN
		SCALE_D := O_LO;
	ELSE
		SCALE_D := (O_HI - O_LO) / UDINT_TO_REAL(DWORD_TO_UDINT(I_HI) - DWORD_TO_UDINT(I_LO)) * UDINT_TO_REAL(LIMIT(DWORD_TO_UDINT(I_LO),DWORD_TO_UDINT(X),DWORD_TO_UDINT(I_HI)) - DWORD_TO_UDINT(I_LO)) + O_LO;
	END_IF;
END_FUNCTION

PROGRAM program0
  VAR
		X :	DWORD;
		I_LO :	DWORD;
		I_HI :	DWORD;
		O_LO :	REAL;
		O_HI :	REAL;
		CEIL5_OUT : REAL;
  END_VAR

  CEIL5_OUT := SCALE_D(X, I_LO, I_HI, O_LO, O_HI);
END_PROGRAM

CONFIGURATION Config0

  RESOURCE Res0 ON PLC
    TASK task0(INTERVAL := T#20ms,PRIORITY := 0);
    PROGRAM instance0 WITH task0 : program0;
  END_RESOURCE
END_CONFIGURATION

(* ---- SCALE_R.ST ---- *)
FUNCTION SCALE_R:REAL
	VAR_INPUT
		X :	REAL;
		I_LO :	REAL;
		I_HI :	REAL;
		O_LO :	REAL;
		O_HI :	REAL;
	END_VAR

	IF I_LO = I_HI THEN
		SCALE_R := O_LO;
	ELSE
		SCALE_R := (O_HI - O_LO) / (I_HI - I_LO) * (LIMIT(I_LO, X, I_HI) - I_LO) + O_LO;
	END_IF;

END_FUNCTION

PROGRAM program0

  	VAR
		X :	REAL;
		I_LO :	REAL;
		I_HI :	REAL;
		O_LO :	REAL;
		O_HI :	REAL;
		CEIL5_OUT : REAL;
  	END_VAR

  	CEIL5_OUT := SCALE_R(X, I_LO, I_HI, O_LO, O_HI);
END_PROGRAM

CONFIGURATION Config0

	RESOURCE Res0 ON PLC
		TASK task0(INTERVAL := T#20ms,PRIORITY := 0);
		PROGRAM instance0 WITH task0 : program0;
	END_RESOURCE

END_CONFIGURATION

(* ---- SCALE_X2.ST ---- *)
FUNCTION SCALE_X2:REAL
	VAR_INPUT
		IN1 :	BOOL;
		IN2 :	BOOL;
		K :	REAL;
		O :	REAL;
		IN1_MIN :	REAL;(*Standard = 0*)
		IN1_MAX :	REAL;(*Standard = 1000*)
		IN2_MIN :	REAL;(*Standard = 0*)
		IN2_MAX :	REAL;(*Standard = 1000*)
	END_VAR

	SCALE_X2 := (SEL(IN1,IN1_MIN, IN1_MAX)+ SEL(IN2,IN2_MIN, IN2_MAX))* k + o;

END_FUNCTION

PROGRAM program0

  	VAR
		IN1 :	BOOL;
		IN2 :	BOOL;
		K :	REAL;
		O :	REAL;
		IN1_MIN :	REAL;(*Standard = 0*)
		IN1_MAX :	REAL;(*Standard = 1000*)
		IN2_MIN :	REAL;(*Standard = 0*)
		IN2_MAX :	REAL;(*Standard = 1000*)
		CEIL5_OUT : REAL;
  	END_VAR

  	CEIL5_OUT := SCALE_X2(IN1, IN2, K, O, IN1_MIN, IN1_MAX, IN2_MIN, IN2_MAX);
END_PROGRAM

CONFIGURATION Config0

	RESOURCE Res0 ON PLC
		TASK task0(INTERVAL := T#20ms,PRIORITY := 0);
		PROGRAM instance0 WITH task0 : program0;
	END_RESOURCE

END_CONFIGURATION

(* ---- SCALE_X4.ST ---- *)
FUNCTION SCALE_X4:REAL
	VAR_INPUT
		IN1 :	BOOL;
		IN2 :	BOOL;
		IN3 :	BOOL;
		IN4 :	BOOL;
		K :	REAL;
		O :	REAL;
		IN1_MIN :	REAL;
		IN1_MAX :	REAL;
		IN2_MIN :	REAL;
		IN2_MAX :	REAL;
		IN3_MIN :	REAL;
		IN3_MAX :	REAL;
		IN4_MIN :	REAL;
		IN4_MAX :	REAL;
	END_VAR
	IF NOT in1 THEN scale_X4 := in1_min; ELSE scale_X4 := in1_max; END_IF;
	IF NOT in2 THEN scale_x4 := scale_x4 + in2_min; ELSE scale_x4 := scale_x4 + in2_max; END_IF;
	IF NOT in3 THEN scale_x4 := scale_x4 + in3_min; ELSE scale_x4 := scale_x4 + in3_max; END_IF;
	IF NOT in4 THEN scale_x4 := scale_x4 + in4_min; ELSE scale_x4 := scale_x4 + in4_max; END_IF;
	scale_X4 := scale_X4 * k + O;
	END_FUNCTION

PROGRAM program0

  	VAR
		IN1 :	BOOL;
		IN2 :	BOOL;
		IN3 :	BOOL;
		IN4 :	BOOL;
		K :	REAL;
		O :	REAL;
		IN1_MIN :	REAL;
		IN1_MAX :	REAL;
		IN2_MIN :	REAL;
		IN2_MAX :	REAL;
		IN3_MIN :	REAL;
		IN3_MAX :	REAL;
		IN4_MIN :	REAL;
		IN4_MAX :	REAL;
		CEIL5_OUT : REAL;
  	END_VAR

  	CEIL5_OUT := SCALE_X4(IN1, IN2, IN3, IN4, K, O, IN1_MIN, IN1_MAX, IN2_MIN, IN2_MAX, IN3_MIN, IN3_MAX, IN4_MIN, IN4_MAX);
END_PROGRAM

CONFIGURATION Config0

	RESOURCE Res0 ON PLC
		TASK task0(INTERVAL := T#20ms,PRIORITY := 0);
		PROGRAM instance0 WITH task0 : program0;
	END_RESOURCE

END_CONFIGURATION

(* ---- SCALE_X8.ST ---- *)
FUNCTION SCALE_X8:REAL

	VAR_INPUT
		IN1 :	BOOL;
		IN2 :	BOOL;
		IN3 :	BOOL;
		IN4 :	BOOL;
		IN5 :	BOOL;
		IN6 :	BOOL;
		IN7 :	BOOL;
		IN8 :	BOOL;
		K :	REAL;
		O :	REAL;
		IN1_MIN :	REAL;
		IN1_MAX :	REAL;
		IN2_MIN :	REAL;
		IN2_MAX :	REAL;
		IN3_MIN :	REAL;
		IN3_MAX :	REAL;
		IN4_MIN :	REAL;
		IN4_MAX :	REAL;
		IN5_MIN :	REAL;
		IN5_MAX :	REAL;
		IN6_MIN :	REAL;
		IN6_MAX :	REAL;
		IN7_MIN :	REAL;
		IN7_MAX :	REAL;
		IN8_MIN :	REAL;
		IN8_MAX :	REAL;
	END_VAR

	SCALE_X8 := (SEL(IN1,IN1_MIN, IN1_MAX)+ SEL(IN2,IN2_MIN, IN2_MAX)+SEL(IN3,IN3_MIN, IN3_MAX)+ SEL(IN4,IN4_MIN, IN4_MAX)
					+SEL(IN5,IN5_MIN, IN5_MAX)+ SEL(IN6,IN6_MIN, IN6_MAX)+SEL(IN7,IN7_MIN, IN7_MAX)+ SEL(IN8,IN8_MIN, IN8_MAX))*k + o;

END_FUNCTION

PROGRAM program0

  	VAR
		IN1 :	BOOL;
		IN2 :	BOOL;
		IN3 :	BOOL;
		IN4 :	BOOL;
		IN5 :	BOOL;
		IN6 :	BOOL;
		IN7 :	BOOL;
		IN8 :	BOOL;
		K :	REAL;
		O :	REAL;
		IN1_MIN :	REAL;
		IN1_MAX :	REAL;
		IN2_MIN :	REAL;
		IN2_MAX :	REAL;
		IN3_MIN :	REAL;
		IN3_MAX :	REAL;
		IN4_MIN :	REAL;
		IN4_MAX :	REAL;
		IN5_MIN :	REAL;
		IN5_MAX :	REAL;
		IN6_MIN :	REAL;
		IN6_MAX :	REAL;
		IN7_MIN :	REAL;
		IN7_MAX :	REAL;
		IN8_MIN :	REAL;
		IN8_MAX :	REAL;
		CEIL5_OUT : REAL;
  	END_VAR

  	CEIL5_OUT := SCALE_X8(IN1, IN2, IN3, IN4, IN5, IN6, IN7, IN8, K, O, IN1_MIN, IN1_MAX, IN2_MIN, IN2_MAX, IN3_MIN, IN3_MAX, IN4_MIN, IN4_MAX, IN5_MIN, IN5_MAX, IN6_MIN, IN6_MAX, IN7_MIN, IN7_MAX, IN8_MIN, IN8_MAX);
END_PROGRAM

CONFIGURATION Config0

	RESOURCE Res0 ON PLC
		TASK task0(INTERVAL := T#20ms,PRIORITY := 0);
		PROGRAM instance0 WITH task0 : program0;
	END_RESOURCE

END_CONFIGURATION

(* ---- SDD.ST ---- *)
FUNCTION SDD:REAL

	VAR_INPUT
		T :	REAL;
		ICE :	BOOL;
	END_VAR

	IF ice THEN
		SDD := 611.153 * EXP(22.4433 * T / (272.186 + T));
	ELSE
		SDD := 611.213 * EXP(17.5043 * T / (241.2 + T));
	END_IF;

END_FUNCTION

PROGRAM program0
  VAR
    T :	REAL;
	ICE :	BOOL;
    CEIL5_OUT : REAL;
  END_VAR

  CEIL5_OUT := SDD(T, ICE);
END_PROGRAM

CONFIGURATION Config0

  RESOURCE Res0 ON PLC
    TASK task0(INTERVAL := T#20ms,PRIORITY := 0);
    PROGRAM instance0 WITH task0 : program0;
  END_RESOURCE
END_CONFIGURATION

(* ---- SDD_NH3.ST ---- *)
FUNCTION SDD_NH3:REAL

	VAR_INPUT
		T :	REAL;
	END_VAR

	IF T < -33.65 THEN
		SDD_NH3 := EXP(7.3396511649 - ( 1166.7498002 / ( T + 192.37 )));
	ELSE
		SDD_NH3 := EXP(11.210964456 - ( 2564.9140075 / ( T + 262.741 )));
	END_IF;

END_FUNCTION

PROGRAM program0
  VAR
    T :	REAL;
    CEIL5_OUT : REAL;
  END_VAR

  CEIL5_OUT := SDD_NH3(T);
END_PROGRAM

CONFIGURATION Config0

  RESOURCE Res0 ON PLC
    TASK task0(INTERVAL := T#20ms,PRIORITY := 0);
    PROGRAM instance0 WITH task0 : program0;
  END_RESOURCE
END_CONFIGURATION

(* ---- SDT_NH3.ST ---- *)
FUNCTION SDT_NH3:REAL

	VAR_INPUT
		P :	REAL;
	END_VAR

	IF P < 1.0E-3 THEN
		SDT_NH3 := -110.0;
	ELSIF P < 1.0 THEN
		SDT_NH3 := 506.713 / (3.18757 - LOG(P)) - 192.37 ;
	ELSE
		SDT_NH3 := 1113.928 / (4.86886 - LOG(P)) - 262.71 ;
	END_IF;

END_FUNCTION

PROGRAM program0
  VAR
    P :	REAL;
    CEIL5_OUT : REAL;
  END_VAR

  CEIL5_OUT := SDT_NH3(P);
END_PROGRAM

CONFIGURATION Config0

  RESOURCE Res0 ON PLC
    TASK task0(INTERVAL := T#20ms,PRIORITY := 0);
    PROGRAM instance0 WITH task0 : program0;
  END_RESOURCE
END_CONFIGURATION

(* ---- SECOND.ST ---- *)
FUNCTION SECOND:REAL

	VAR_INPUT
		ITOD :	UDINT;
	END_VAR

	second := UDINT_TO_REAL(itod MOD UDINT#60000) / REAL#1000.00;

END_FUNCTION

PROGRAM program0
  VAR
    ITOD :	UDINT;
    CEIL5_OUT : REAL;
  END_VAR

  CEIL5_OUT := SECOND(ITOD);
END_PROGRAM

CONFIGURATION Config0

	RESOURCE Res0 ON PLC
		TASK task0(INTERVAL := T#20ms,PRIORITY := 0);
		PROGRAM instance0 WITH task0 : program0;
	END_RESOURCE

END_CONFIGURATION

(* ---- SECOND_OF_DT.ST ---- *)
FUNCTION SECOND_OF_DT:INT

	VAR_INPUT
		XDT :	UDINT;
	END_VAR

	SECOND_OF_DT := UDINT_TO_INT(XDT MOD UDINT#60);
END_FUNCTION

PROGRAM program0
  VAR
    LocalVar0 : UDINT;
	LocalOUT  : INT;
  END_VAR
  	LocalOUT := SECOND_OF_DT(LocalVar0);
END_PROGRAM

CONFIGURATION Config0
  RESOURCE Res0 ON PLC
    TASK task0(INTERVAL := T#20ms,PRIORITY := 0);
    PROGRAM instance0 WITH task0 : program0;
  END_RESOURCE
END_CONFIGURATION

(* ---- SECOND_TO_TIME.ST ---- *)
FUNCTION _REAL_TO_UDINT:UDINT
	VAR_INPUT
		X :	REAL;
	END_VAR

	IF REAL_TO_UDINT(0.5) = UDINT#1 THEN
		_REAL_TO_UDINT := REAL_TO_UDINT(x);
	ELSIF X > 0.0 THEN
		_REAL_TO_UDINT := REAL_TO_UDINT(x+0.5);
	ELSIF X < 0.0 THEN
		_REAL_TO_UDINT := REAL_TO_UDINT(x-0.5);
	ELSE
		_REAL_TO_UDINT := UDINT#0;
	END_IF;
END_FUNCTION

FUNCTION SECOND_TO_TIME:TIME

	VAR_INPUT
		IN :	REAL;
	END_VAR

	second_to_time := UDINT_TO_TIME(_REAL_TO_UDINT(IN * 1000.0));

END_FUNCTION

PROGRAM program0

	VAR
		IN :	REAL;
		CEIL5_OUT : TIME;
	END_VAR

	CEIL5_OUT := SECOND_TO_TIME(IN);

END_PROGRAM

CONFIGURATION Config0

	RESOURCE Res0 ON PLC
		TASK task0(INTERVAL := T#20ms,PRIORITY := 0);
		PROGRAM instance0 WITH task0 : program0;
	END_RESOURCE

END_CONFIGURATION

(* ---- SENSOR_INT.ST ---- *)
FUNCTION SENSOR_INT:REAL

	VAR_INPUT
		VOLTAGE :	REAL;
		CURRENT :	REAL;
		RP :	REAL;
		_RS :	REAL;
	END_VAR

	VAR
		RG :	REAL;
	END_VAR

	IF current <> 0.0 THEN
		RG := voltage / current;
		SENSOR_INT := RP * ( RG - _RS) / ( RP + _RS - RG);
	END_IF;

END_FUNCTION

PROGRAM program0

	VAR
		VOLTAGE :	REAL;
		CURRENT :	REAL;
		RP :	REAL;
		_RS :	REAL;
		CEIL5_OUT : REAL;
	END_VAR

	CEIL5_OUT := SENSOR_INT(VOLTAGE, CURRENT, RP, _RS);

END_PROGRAM

CONFIGURATION Config0

	RESOURCE Res0 ON PLC
		TASK task0(INTERVAL := T#20ms,PRIORITY := 0);
		PROGRAM instance0 WITH task0 : program0;
	END_RESOURCE

END_CONFIGURATION

(* ---- SET_DATE.ST ---- *)
FUNCTION _INT_TO_UDINT:UDINT
	VAR_INPUT
		IN :	INT;
	END_VAR

	_INT_TO_UDINT := DINT_TO_UDINT(INT_TO_DINT(IN));
END_FUNCTION

FUNCTION SET_DATE:UDINT

	VAR_INPUT
		YEAR :	INT;
		MONTH :	INT;
		DAY :	INT;
	END_VAR

	VAR
		count :	INT;
	END_VAR

	IF month > 2 THEN
		count := (month - 1) * 30;
		IF month > 7 THEN
			count := count + DWORD_TO_INT(SHR(DINT_TO_DWORD(INT_TO_DINT(month) - INT_TO_DINT(3)),1));
		ELSE
			count := count + DWORD_TO_INT(SHR(DINT_TO_DWORD(INT_TO_DINT(month) - INT_TO_DINT(4)),1));
		END_IF;
		IF SHL(INT_TO_WORD(year),14) = WORD#0 THEN
			count := count + 1;
		END_IF;
	ELSE
		count := (month - 1) * 31;
	END_IF;
	SET_DATE := (_INT_TO_UDINT(count + day - 1) + DWORD_TO_UDINT(SHR(UDINT_TO_DWORD(_INT_TO_UDINT(year) * UDINT#1461 - UDINT#2878169), 2))) * UDINT#86400;

END_FUNCTION

PROGRAM program0
  VAR
	YEAR :	INT;
	MONTH :	INT;
	DAY :	INT;
    CEIL5_OUT : UDINT;
  END_VAR

  CEIL5_OUT := SET_DATE(YEAR, MONTH, DAY);
END_PROGRAM

CONFIGURATION Config0

  RESOURCE Res0 ON PLC
    TASK task0(INTERVAL := T#20ms,PRIORITY := 0);
    PROGRAM instance0 WITH task0 : program0;
  END_RESOURCE
END_CONFIGURATION

(* ---- SET_DT.ST ---- *)
FUNCTION _INT_TO_UDINT:UDINT
	VAR_INPUT
		IN :	INT;
	END_VAR

	_INT_TO_UDINT := DINT_TO_UDINT(INT_TO_DINT(IN));
END_FUNCTION

FUNCTION SET_DATE:UDINT

	VAR_INPUT
		YEAR :	INT;
		MONTH :	INT;
		DAY :	INT;
	END_VAR

	VAR
		count :	INT;
	END_VAR

	IF month > 2 THEN
		count := (month - 1) * 30;
		IF month > 7 THEN
			count := count + DWORD_TO_INT(SHR(DINT_TO_DWORD(INT_TO_DINT(month) - INT_TO_DINT(3)),1));
		ELSE
			count := count + DWORD_TO_INT(SHR(DINT_TO_DWORD(INT_TO_DINT(month) - INT_TO_DINT(4)),1));
		END_IF;
		IF SHL(INT_TO_WORD(year),14) = WORD#0 THEN
			count := count + 1;
		END_IF;
	ELSE
		count := (month - 1) * 31;
	END_IF;
	SET_DATE := (_INT_TO_UDINT(count + day - 1) + DWORD_TO_UDINT(SHR(UDINT_TO_DWORD(_INT_TO_UDINT(year) * UDINT#1461 - UDINT#2878169), 2))) * UDINT#86400;

END_FUNCTION

FUNCTION SET_DT:UDINT
	VAR_INPUT
		YEAR :	INT;
		MONTH :	INT;
		DAY :	INT;
		HOUR :	INT;
		MINUTE :	INT;
		SECOND :	INT;
	END_VAR

	SET_DT := SET_DATE(YEAR, MONTH, DAY) + _INT_TO_UDINT(SECOND) + _INT_TO_UDINT(MINUTE) * UDINT#60 + _INT_TO_UDINT(HOUR) * UDINT#3600;
END_FUNCTION

PROGRAM program0

	VAR
		YEAR :	INT;
		MONTH :	INT;
		DAY :	INT;
		HOUR :	INT;
		MINUTE :	INT;
		SECOND :	INT;
		CEIL5_OUT : UDINT;
	END_VAR

	CEIL5_OUT := SET_DT(YEAR, MONTH, DAY, HOUR, MINUTE, SECOND);

END_PROGRAM

CONFIGURATION Config0

	RESOURCE Res0 ON PLC
		TASK task0(INTERVAL := T#20ms,PRIORITY := 0);
		PROGRAM instance0 WITH task0 : program0;
	END_RESOURCE

END_CONFIGURATION

(* ---- SET_TOD.ST ---- *)
FUNCTION _REAL_TO_UDINT:UDINT

	VAR_INPUT
		X :	REAL;
	END_VAR

	IF REAL_TO_UDINT(0.5) = UDINT#1 THEN
		_REAL_TO_UDINT := REAL_TO_UDINT(x);
	ELSIF X > 0.0 THEN
		_REAL_TO_UDINT := REAL_TO_UDINT(x+0.5);
	ELSIF X < 0.0 THEN
		_REAL_TO_UDINT := REAL_TO_UDINT(x-0.5);
	ELSE
		_REAL_TO_UDINT := UDINT#0;
	END_IF;

END_FUNCTION

FUNCTION _INT_TO_UDINT:UDINT

	VAR_INPUT
		IN :	INT;
	END_VAR

	_INT_TO_UDINT := DINT_TO_UDINT(INT_TO_DINT(IN));

END_FUNCTION

FUNCTION SET_TOD:UDINT

	VAR_INPUT
		HOUR :	INT;
		MINUTE :	INT;
		SECOND :	REAL;
	END_VAR

	set_Tod := _REAL_TO_UDINT(second * 1000.0) + _INT_TO_UDINT(minute) * UDINT#60000 + _INT_TO_UDINT(hour) * UDINT#3600000;

END_FUNCTION

PROGRAM program0

	VAR
		HOUR :	INT;
		MINUTE :	INT;
		SECOND :	REAL;
		CEIL5_OUT : UDINT;
	END_VAR

	CEIL5_OUT := SET_TOD(HOUR, MINUTE, SECOND);

END_PROGRAM

CONFIGURATION Config0

	RESOURCE Res0 ON PLC
		TASK task0(INTERVAL := T#20ms,PRIORITY := 0);
		PROGRAM instance0 WITH task0 : program0;
	END_RESOURCE

END_CONFIGURATION

(* ---- SETUP_EXTENDED_ASCII.ST ---- *)
FUNCTION SETUP_EXTENDED_ASCII:BOOL

	VAR_INPUT
		X :	BOOL;
	END_VAR

	SETUP_EXTENDED_ASCII := X OR TRUE;
END_FUNCTION

PROGRAM program0
  VAR
	X :	BOOL;
    CEIL5_OUT : BOOL;
  END_VAR

  CEIL5_OUT := SETUP_EXTENDED_ASCII(X);
END_PROGRAM

CONFIGURATION Config0

  RESOURCE Res0 ON PLC
    TASK task0(INTERVAL := T#20ms,PRIORITY := 0);
    PROGRAM instance0 WITH task0 : program0;
  END_RESOURCE
END_CONFIGURATION

(* ---- SGN.ST ---- *)
FUNCTION SGN : INT
  VAR_INPUT
    x : REAL;
  END_VAR

  IF X > 0.0 THEN
  	sgn := 1;
  ELSIF X < 0.0 THEN
  	sgn := -1;
  ELSE
  	sgn := 0;
  END_IF;
END_FUNCTION

PROGRAM program0
  VAR
    LocalVar0 : REAL;
    LocalVar1 : INT;
    CEIL5_OUT : INT;
  END_VAR

  CEIL5_OUT := SGN(LocalVar0);
  LocalVar1 := CEIL5_OUT;
END_PROGRAM

CONFIGURATION Config0

  RESOURCE Res0 ON PLC
    TASK task0(INTERVAL := T#20ms,PRIORITY := 0);
    PROGRAM instance0 WITH task0 : program0;
  END_RESOURCE
END_CONFIGURATION

(* ---- SHL1.ST ---- *)
FUNCTION SHL1:DWORD

	VAR_INPUT
		IN :	DWORD;
		N :	INT;
	END_VAR

	SHL1 := SHR(DWORD#16#FF_FF_FF_FF,32-N) OR SHL(IN,N);

END_FUNCTION

PROGRAM program0

	VAR
		IN :	DWORD;
		N :	INT;
		CEIL5_OUT : DWORD;
	END_VAR

  	CEIL5_OUT := SHL1(IN, N);

END_PROGRAM

CONFIGURATION Config0

	RESOURCE Res0 ON PLC
		TASK task0(INTERVAL := T#20ms,PRIORITY := 0);
		PROGRAM instance0 WITH task0 : program0;
	END_RESOURCE

END_CONFIGURATION

(* ---- SHR1.ST ---- *)
FUNCTION SHR1:DWORD

	VAR_INPUT
		IN :	DWORD;
		N :	INT;
	END_VAR

	SHR1 := SHL(DWORD#16#FF_FF_FF_FF,32-N) OR SHR(IN,N);

END_FUNCTION

PROGRAM program0

	VAR
		IN : DWORD;
		N :	INT;
		CEIL5_OUT : DWORD;
	END_VAR

	CEIL5_OUT := SHR1(IN, N);

END_PROGRAM

CONFIGURATION Config0

	RESOURCE Res0 ON PLC
		TASK task0(INTERVAL := T#20ms,PRIORITY := 0);
		PROGRAM instance0 WITH task0 : program0;
	END_RESOURCE

END_CONFIGURATION

(* ---- SIGMOID.ST ---- *)
FUNCTION SIGMOID:REAL

	VAR_INPUT
		X :	REAL;
	END_VAR

	IF X > 20.0 THEN
		SIGMOID := 1.0;
	ELSIF x < -85.0 THEN
		SIGMOID := 0.0;
	ELSE
		SIGMOID := 1.0 / (1.0 + EXP(-X));
	END_IF;

END_FUNCTION

PROGRAM program0

	VAR
		X :	REAL;
		CEIL5_OUT : REAL;
	END_VAR

	CEIL5_OUT := SIGMOID(X);

END_PROGRAM

CONFIGURATION Config0

	RESOURCE Res0 ON PLC
		TASK task0(INTERVAL := T#20ms,PRIORITY := 0);
		PROGRAM instance0 WITH task0 : program0;
	END_RESOURCE

END_CONFIGURATION

(* ---- SIGN_I.ST ---- *)
FUNCTION BIT_OF_DWORD : BOOL

	VAR_INPUT
		IN : DWORD;
		N : INT;
	END_VAR

	BIT_OF_DWORD := (SHR(in,N) AND 16#00000001) > 0;

END_FUNCTION

FUNCTION SIGN_I:BOOL

	VAR_INPUT
		IN :	DINT;
	END_VAR

	sign_I := BIT_OF_DWORD(DINT_TO_DWORD(in),31);

END_FUNCTION

PROGRAM program0

	VAR
		IN :	DINT;
		CEIL5_OUT : BOOL;
	END_VAR

	CEIL5_OUT := SIGN_I(IN);

END_PROGRAM

CONFIGURATION Config0

	RESOURCE Res0 ON PLC
		TASK task0(INTERVAL := T#20ms,PRIORITY := 0);
		PROGRAM instance0 WITH task0 : program0;
	END_RESOURCE

END_CONFIGURATION

(* ---- SIGN_R.ST ---- *)
FUNCTION SIGN_R : BOOL
  VAR_INPUT
    IN : REAL;
  END_VAR

  SIGN_R := in < 0.0;
END_FUNCTION

PROGRAM program0
  VAR
    LocalVar0 : REAL;
    CEIL5_OUT : BOOL;
  END_VAR

  CEIL5_OUT := SIGN_R(LocalVar0);
END_PROGRAM

CONFIGURATION Config0

  RESOURCE Res0 ON PLC
    TASK task0(INTERVAL := T#20ms,PRIORITY := 0);
    PROGRAM instance0 WITH task0 : program0;
  END_RESOURCE
END_CONFIGURATION

(* ---- SINC.ST ---- *)
FUNCTION SINC:REAL

	VAR_INPUT
		X :	REAL;
	END_VAR

	IF X = 0.0 THEN
		SINC := 1.0;
	ELSE
		SINC := SIN(x) / x;
	END_IF;

END_FUNCTION

PROGRAM program0

	VAR
		X :	REAL;
		CEIL5_OUT : REAL;
	END_VAR

  	CEIL5_OUT := SINC(X);

END_PROGRAM

CONFIGURATION Config0

	RESOURCE Res0 ON PLC
		TASK task0(INTERVAL := T#20ms,PRIORITY := 0);
		PROGRAM instance0 WITH task0 : program0;
	END_RESOURCE

END_CONFIGURATION

(* ---- SINH.ST ---- *)
FUNCTION SINH:REAL
	VAR_INPUT
		X :	REAL;
	END_VAR

	IF ABS(x) < 2.0E-3 THEN
		SINH := X;
	ELSE
		SINH := (EXP(x) - EXP(-x)) * 0.5;
	END_IF;
END_FUNCTION

PROGRAM program0
  VAR
    LocalVar0 : REAL;
    CEIL5_OUT : REAL;
  END_VAR

  CEIL5_OUT := SINH(LocalVar0);
END_PROGRAM

CONFIGURATION Config0

  RESOURCE Res0 ON PLC
    TASK task0(INTERVAL := T#20ms,PRIORITY := 0);
    PROGRAM instance0 WITH task0 : program0;
  END_RESOURCE
END_CONFIGURATION

(* ---- SPHERE_V.ST ---- *)
FUNCTION SPHERE_V:REAL

	VAR_INPUT
		RX :	REAL;
	END_VAR

	sphere_V := 4.188790205 * Rx * RX * RX;

END_FUNCTION

PROGRAM program0

	VAR
		RX :	REAL;
		CEIL5_OUT : REAL;
	END_VAR

	CEIL5_OUT := SPHERE_V(RX);

END_PROGRAM

CONFIGURATION Config0

	RESOURCE Res0 ON PLC
		TASK task0(INTERVAL := T#20ms,PRIORITY := 0);
		PROGRAM instance0 WITH task0 : program0;
	END_RESOURCE

END_CONFIGURATION

(* ---- SQRTN.ST ---- *)
FUNCTION SQRTN:REAL

	VAR_INPUT
		X :	REAL;
		N :	INT;
	END_VAR

	IF N > 0 THEN
		SQRTN := EXP(LN(x) / INT_TO_REAL(n));
	ELSE
		SQRTN := 0.0;
	END_IF;

END_FUNCTION

PROGRAM program0
	VAR
		LocalVar0 : REAL;
		LocalVar1 : INT;
		LocalOUT  : REAL;
	END_VAR

 	LocalOUT := SQRTN(LocalVar0, LocalVar1);

END_PROGRAM

CONFIGURATION Config0

	RESOURCE Res0 ON PLC
		TASK task0(INTERVAL := T#20ms,PRIORITY := 0);
		PROGRAM instance0 WITH task0 : program0;
	END_RESOURCE

END_CONFIGURATION

(* ---- STAIR.ST ---- *)
FUNCTION _REAL_TO_DINT:DINT
	VAR_INPUT
		X :	REAL;
	END_VAR

	IF REAL_TO_DINT(0.5) = DINT#1 THEN
		_REAL_TO_DINT := REAL_TO_DINT(x);
		RETURN;
	END_IF;

	IF X > 0.0 THEN
		_REAL_TO_DINT := REAL_TO_DINT(x+0.5);
	ELSIF X < 0.0 THEN
		_REAL_TO_DINT := REAL_TO_DINT(x-0.5);
	ELSE
		_REAL_TO_DINT := DINT#0;
	END_IF;

END_FUNCTION

FUNCTION STAIR:REAL

	VAR_INPUT
		X :	REAL;
		D :	REAL;
	END_VAR

	IF D > 0.0 THEN
		STAIR := DINT_TO_REAL(_REAL_TO_DINT(X / D)) * D;
	ELSE
		STAIR := X;
	END_IF;

END_FUNCTION

PROGRAM program0

	VAR
		X :	REAL;
		D :	REAL;
		CEIL5_OUT : REAL;
	END_VAR

	CEIL5_OUT := STAIR(X, D);

END_PROGRAM

CONFIGURATION Config0

	RESOURCE Res0 ON PLC
		TASK task0(INTERVAL := T#20ms,PRIORITY := 0);
		PROGRAM instance0 WITH task0 : program0;
	END_RESOURCE

END_CONFIGURATION

(* ---- SUN_MIDDAY.ST ---- *)
FUNCTION _REAL_TO_UDINT:UDINT
	VAR_INPUT
		X :	REAL;
	END_VAR

	IF REAL_TO_UDINT(0.5) = UDINT#1 THEN
		_REAL_TO_UDINT := REAL_TO_UDINT(x);
	ELSIF X > 0.0 THEN
		_REAL_TO_UDINT := REAL_TO_UDINT(x+0.5);
	ELSIF X < 0.0 THEN
		_REAL_TO_UDINT := REAL_TO_UDINT(x-0.5);
	ELSE
		_REAL_TO_UDINT := UDINT#0;
	END_IF;

END_FUNCTION

FUNCTION HOUR_TO_TOD:UDINT

	VAR_INPUT
		IN :	REAL;
	END_VAR

	hour_to_tod := _REAL_TO_UDINT(IN * 3600000.00);

END_FUNCTION

FUNCTION DAY_OF_YEAR:INT
	VAR_INPUT
		IDATE :	DATE;
	END_VAR

	DAY_OF_YEAR := UDINT_TO_INT((DATE_TO_UDINT(idate) / UDINT#86400) MOD UDINT#1461);
	IF DAY_OF_YEAR > 729 THEN
		IF DAY_OF_YEAR > 1095 THEN DAY_OF_YEAR := DAY_OF_YEAR - 1095; ELSE DAY_OF_YEAR := DAY_OF_YEAR - 729; END_IF;
	ELSIF DAY_OF_YEAR > 364 THEN
		DAY_OF_YEAR := DAY_OF_YEAR - 364;
	ELSE
		DAY_OF_YEAR := DAY_OF_YEAR + 1;
	END_IF;
END_FUNCTION

FUNCTION SUN_MIDDAY:UDINT

	VAR_INPUT
		LON :	REAL;
		UTC :	DATE;
	END_VAR

	VAR
		T :	REAL;
		OFFSET :	REAL;
	END_VAR

	T := INT_TO_REAL(DAY_OF_YEAR(utc));
	OFFSET := -0.1752 * SIN(0.033430 * T + 0.5474) - 0.1340 * SIN(0.018234 * T - 0.1939);
	SUN_MIDDAY := HOUR_TO_TOD(12.0 - OFFSET - lon * 0.0666666666666);

END_FUNCTION

PROGRAM program0

	VAR
		LON :	REAL;
		UTC :	DATE;
		CEIL5_OUT : UDINT;
	END_VAR

	CEIL5_OUT := SUN_MIDDAY(LON, UTC);

END_PROGRAM

CONFIGURATION Config0

	RESOURCE Res0 ON PLC
		TASK task0(INTERVAL := T#20ms,PRIORITY := 0);
		PROGRAM instance0 WITH task0 : program0;
	END_RESOURCE

END_CONFIGURATION

(* ---- SWAP_BYTE.ST ---- *)
FUNCTION SWAP_BYTE:WORD

	VAR_INPUT
		IN :	WORD;
	END_VAR

	Swap_Byte := ROL(in,8);

END_FUNCTION

PROGRAM program0

	VAR
		IN :	WORD;
		CEIL5_OUT : WORD;
	END_VAR

	CEIL5_OUT := SWAP_BYTE(IN);

END_PROGRAM

CONFIGURATION Config0

	RESOURCE Res0 ON PLC
		TASK task0(INTERVAL := T#20ms,PRIORITY := 0);
		PROGRAM instance0 WITH task0 : program0;
	END_RESOURCE

END_CONFIGURATION

(* ---- SWAP_BYTE2.ST ---- *)
FUNCTION SWAP_BYTE2:DWORD

	VAR_INPUT
		INPUT :	DWORD;
	END_VAR

	Swap_Byte2 := (ROR(INPUT,8) AND DWORD#16#FF00FF00) OR (ROL(INPUT,8) AND DWORD#16#00FF00FF);

END_FUNCTION

PROGRAM program0

	VAR
		IN :	DWORD;
		CEIL5_OUT : DWORD;
	END_VAR

	CEIL5_OUT := SWAP_BYTE2(IN);

END_PROGRAM

CONFIGURATION Config0

	RESOURCE Res0 ON PLC
		TASK task0(INTERVAL := T#20ms,PRIORITY := 0);
		PROGRAM instance0 WITH task0 : program0;
	END_RESOURCE

END_CONFIGURATION

(* ---- TANC.ST ---- *)
FUNCTION TANC:REAL

	VAR_INPUT
		X :	REAL;
	END_VAR

	IF X = 0.0 THEN
		TANC := 1.0;
	ELSE
		TANC := TAN(x) / x;
	END_IF;

END_FUNCTION

PROGRAM program0

	VAR
		X :	REAL;
		CEIL5_OUT : REAL;
	END_VAR

	CEIL5_OUT := TANC(X);

END_PROGRAM

CONFIGURATION Config0

	RESOURCE Res0 ON PLC
		TASK task0(INTERVAL := T#20ms,PRIORITY := 0);
		PROGRAM instance0 WITH task0 : program0;
	END_RESOURCE

END_CONFIGURATION

(* ---- TANH.ST ---- *)
FUNCTION TANH:REAL

	VAR_INPUT
		X :	REAL;
	END_VAR

	IF X > 20.0 THEN
		TANH := 1.0;
	ELSIF X < -20.0 THEN
		TANH := -1.0;
	ELSE
		TANH := 1.0 - 2.0 / (EXP(2.0 * x) + 1.0);
	END_IF;

END_FUNCTION

PROGRAM program0

	VAR
		X :	REAL;
		CEIL5_OUT : REAL;
	END_VAR

	CEIL5_OUT := TANH(X);

END_PROGRAM

CONFIGURATION Config0

	RESOURCE Res0 ON PLC
		TASK task0(INTERVAL := T#20ms,PRIORITY := 0);
		PROGRAM instance0 WITH task0 : program0;
	END_RESOURCE

END_CONFIGURATION

(* ---- TANK_VOL1.ST ---- *)
FUNCTION CIRCLE_SEG:REAL
	VAR_INPUT
		RX :	REAL;
		HX :	REAL;
	END_VAR

	IF RX > 0.0 THEN
		CIRCLE_SEG := 2.0 * ACOS(1.0 - LIMIT(0.0, HX / RX, 2.0));
		CIRCLE_SEG := (CIRCLE_SEG - SIN(CIRCLE_SEG)) * RX * RX * 0.5;
	END_IF;
END_FUNCTION

FUNCTION TANK_VOL1:REAL

	VAR_INPUT
		TR :	REAL;
		TL :	REAL;
		H :	REAL;
	END_VAR

	TANK_VOL1 := CIRCLE_SEG(TR, H) * TL;

END_FUNCTION

PROGRAM program0
  VAR
    TR :	REAL;
	TL :	REAL;
	H :	REAL;
    CEIL5_OUT : REAL;
  END_VAR

  CEIL5_OUT := TANK_VOL1(TR, TL, H);
END_PROGRAM

CONFIGURATION Config0

  RESOURCE Res0 ON PLC
    TASK task0(INTERVAL := T#20ms,PRIORITY := 0);
    PROGRAM instance0 WITH task0 : program0;
  END_RESOURCE
END_CONFIGURATION

(* ---- TANK_VOL2.ST ---- *)
FUNCTION TANK_VOL2:REAL

	VAR_INPUT
		TR :	REAL;
		H :	REAL;
	END_VAR

	TANK_VOL2 := 3.14159265358979323846264338327950288 * H * H * (TR - H / 3.0);

END_FUNCTION

PROGRAM program0
  VAR
    TR :	REAL;
	H :	REAL;
    CEIL5_OUT : REAL;
  END_VAR

  CEIL5_OUT := TANK_VOL2(TR, H);
END_PROGRAM

CONFIGURATION Config0

  RESOURCE Res0 ON PLC
    TASK task0(INTERVAL := T#20ms,PRIORITY := 0);
    PROGRAM instance0 WITH task0 : program0;
  END_RESOURCE
END_CONFIGURATION

(* ---- TEMP_NI.ST ---- *)
FUNCTION TEMP_NI:REAL
	VAR_INPUT
		RES :	REAL;
		R0 :	REAL;
	END_VAR

	TEMP_NI := (SQRT(0.30085225 - 2.66E-3 * (R0 - Res)) - 0.5485) * 751.8796992;
END_FUNCTION

PROGRAM program0
  	VAR
		RES :	REAL;
		R0 :	REAL;
    	CEIL5_OUT : REAL;
  	END_VAR

  	CEIL5_OUT := TEMP_NI(RES, R0);
END_PROGRAM

CONFIGURATION Config0
	RESOURCE Res0 ON PLC
		TASK task0(INTERVAL := T#20ms,PRIORITY := 0);
		PROGRAM instance0 WITH task0 : program0;
	END_RESOURCE
END_CONFIGURATION

(* ---- TEMP_NTC.ST ---- *)
FUNCTION TEMP_NTC:REAL

VAR_INPUT
	RES :	REAL;
	RN :	REAL;
	B :	REAL;
END_VAR

IF res > 0.0 THEN
	TEMP_NTC := B * 298.15 / (B + LN(RES / RN) * 298.15) -273.15;
END_IF;

END_FUNCTION

PROGRAM program0
  	VAR
		RES :	REAL;
		RN :	REAL;
		B :	REAL;
    	CEIL5_OUT : REAL;
  	END_VAR

  	CEIL5_OUT := TEMP_NTC(RES, RN, B);
END_PROGRAM

CONFIGURATION Config0
	RESOURCE Res0 ON PLC
		TASK task0(INTERVAL := T#20ms,PRIORITY := 0);
		PROGRAM instance0 WITH task0 : program0;
	END_RESOURCE
END_CONFIGURATION

(* ---- TEMP_PT.ST ---- *)
FUNCTION RES_PT:REAL
	VAR_INPUT
		T :	REAL;
		R0 :	REAL;
	END_VAR

	VAR
		T2 :	REAL;
	END_VAR

	T2 := T * T;

	IF T >= 0.0 THEN
		RES_PT := R0 * ( 1.0 + 3.90802E-3 * T + -5.802E-7 * T2);
	ELSE
		RES_PT := R0 * ( 1.0 + 3.90802E-3 * T + -5.802E-7 * T2 + -4.27350E-12 * (T - 100.0) * T2 * T);
	END_IF;

END_FUNCTION

FUNCTION TEMP_PT:REAL

	VAR_INPUT
		RES :	REAL;
		R0 :	REAL;
	END_VAR

	VAR
		step_var :	REAL := REAL#50.0;
		X :	REAL;
		Y :	REAL;
		t1 :	REAL;
	END_VAR

	X := 3.9083E-3 * R0;
	Y := -5.775E-7 * R0;
	IF Res >= R0 THEN
		t1 := X * X - 4.0 * Y * (R0 - Res);
		IF t1 < 0.0 THEN
			TEMP_PT := 10000.0;
		ELSE
			TEMP_PT := (-X + SQRT(t1)) / (2.0 * Y);
		END_IF;
	ELSE
		TEMP_PT := -100.0;
		WHILE step_var > 0.01 DO
			IF RES_PT(TEMP_PT, R0) < res THEN TEMP_PT := TEMP_PT + step_var; ELSE TEMP_PT := TEMP_PT - step_var; END_IF;
			step_var := step_var * 0.5;
		END_WHILE;
	END_IF;
END_FUNCTION

PROGRAM program0
	VAR
		RES :	REAL;
		R0 :	REAL;
		CEIL5_OUT : REAL;
	END_VAR

	CEIL5_OUT := TEMP_PT(RES, R0);
END_PROGRAM

CONFIGURATION Config0
	RESOURCE Res0 ON PLC
		TASK task0(INTERVAL := T#20ms,PRIORITY := 0);
		PROGRAM instance0 WITH task0 : program0;
	END_RESOURCE
END_CONFIGURATION

(* ---- TEMP_SI.ST ---- *)
FUNCTION TEMP_SI:REAL
	VAR_INPUT
		RES :	REAL;
		VAR_RS:	REAL;
		TS :	REAL;
	END_VAR

	TEMP_SI := (-7.64E-3 + SQRT(RES/VAR_RS* 6.64E-5 - 0.803E-5)) * 30120.48193 + TS;

END_FUNCTION

PROGRAM program0
  	VAR
		RES :	REAL;
		VAR_RS:	REAL;
		TS :	REAL;
    	CEIL5_OUT : REAL;
  	END_VAR

  	CEIL5_OUT := TEMP_SI(RES, VAR_RS, TS);
END_PROGRAM

CONFIGURATION Config0
	RESOURCE Res0 ON PLC
		TASK task0(INTERVAL := T#20ms,PRIORITY := 0);
		PROGRAM instance0 WITH task0 : program0;
	END_RESOURCE
END_CONFIGURATION

(* ---- TIME_TO_DWORD.ST ---- *)
FUNCTION TIME_TO_DWORD1:DWORD

VAR_INPUT
	X :	TIME;
END_VAR

TIME_TO_DWORD1 := UDINT_TO_DWORD(DINT_TO_UDINT(TIME_TO_DINT(X)));
END_FUNCTION

PROGRAM program0
  VAR
	X :	TIME;
    CEIL5_OUT : DWORD;
  END_VAR

  CEIL5_OUT := TIME_TO_DWORD1(X);
END_PROGRAM

CONFIGURATION Config0

  RESOURCE Res0 ON PLC
    TASK task0(INTERVAL := T#20ms,PRIORITY := 0);
    PROGRAM instance0 WITH task0 : program0;
  END_RESOURCE
END_CONFIGURATION

(* ---- TIME_TO_INT.ST ---- *)
FUNCTION TIME_TO_INT1:INT

VAR_INPUT
	IN :	TIME;
END_VAR

TIME_TO_INT1 := DINT_TO_INT(TIME_TO_DINT(IN));
END_FUNCTION

PROGRAM program0
  VAR
	IN :	TIME;
    CEIL5_OUT : INT;
  END_VAR

  CEIL5_OUT := TIME_TO_INT1(IN);
END_PROGRAM

CONFIGURATION Config0

  RESOURCE Res0 ON PLC
    TASK task0(INTERVAL := T#20ms,PRIORITY := 0);
    PROGRAM instance0 WITH task0 : program0;
  END_RESOURCE
END_CONFIGURATION

(* ---- TIME_TO_REAL.ST ---- *)
FUNCTION TIME_TO_REAL1:REAL

VAR_INPUT
	X :	TIME;
END_VAR

TIME_TO_REAL1 := UDINT_TO_REAL(DINT_TO_UDINT(TIME_TO_DINT(X)));
END_FUNCTION

PROGRAM program0
  VAR
	X :	TIME;
    CEIL5_OUT : REAL;
  END_VAR

  CEIL5_OUT := TIME_TO_REAL1(X);
END_PROGRAM

CONFIGURATION Config0

  RESOURCE Res0 ON PLC
    TASK task0(INTERVAL := T#20ms,PRIORITY := 0);
    PROGRAM instance0 WITH task0 : program0;
  END_RESOURCE
END_CONFIGURATION

(* ---- TIME_TO_TOD.ST ---- *)
FUNCTION TIME_TO_TOD:UDINT

	VAR_INPUT
		IN :	TIME;
	END_VAR

	TIME_TO_TOD := DWORD_TO_UDINT(TIME_TO_DWORD(IN));
END_FUNCTION

PROGRAM program0
  VAR
	IN :	TIME;
    CEIL5_OUT : UDINT;
  END_VAR

  CEIL5_OUT := TIME_TO_TOD(IN);
END_PROGRAM

CONFIGURATION Config0

  RESOURCE Res0 ON PLC
    TASK task0(INTERVAL := T#20ms,PRIORITY := 0);
    PROGRAM instance0 WITH task0 : program0;
  END_RESOURCE
END_CONFIGURATION

(* ---- TIME_TO_UDINT.ST ---- *)
FUNCTION TIME_TO_UDINT2:UDINT
	VAR_INPUT
		X :	TIME;
	END_VAR

	TIME_TO_UDINT2 := DINT_TO_UDINT(TIME_TO_DINT(X));
END_FUNCTION

PROGRAM program0
  VAR
    LocalVar0 : TIME;
    LocalOUT  : UDINT;
  END_VAR

  LocalOUT := TIME_TO_UDINT2(LocalVar0);
END_PROGRAM

CONFIGURATION Config0
    RESOURCE Res0 ON PLC
        TASK task0(INTERVAL := T#20ms,PRIORITY := 0);
        PROGRAM instance0 WITH task0 : program0;
    END_RESOURCE
END_CONFIGURATION

(* ---- TIMECHECK.ST ---- *)
FUNCTION TIMECHECK:BOOL

	VAR_INPUT
		TD :	UDINT;
		START :	UDINT;
		STOP :	UDINT;
	END_VAR

	IF stop < start THEN
		TIMECHECK := start <= TD OR  TD < stop;
	ELSE
		TIMECHECK := start <= TD AND TD < stop;
	END_IF;

END_FUNCTION

PROGRAM program0
  VAR
	TD :	UDINT;
	START :	UDINT;
	STOP :	UDINT;
    CEIL5_OUT : BOOL;
  END_VAR

  CEIL5_OUT := TIMECHECK(TD, START, STOP);
END_PROGRAM

CONFIGURATION Config0

  RESOURCE Res0 ON PLC
    TASK task0(INTERVAL := T#20ms,PRIORITY := 0);
    PROGRAM instance0 WITH task0 : program0;
  END_RESOURCE
END_CONFIGURATION

(* ---- TN_SC_SHADOW_ATTR.ST ---- *)
FUNCTION TN_SC_SHADOW_ATTR:BYTE

	VAR_INPUT
		Iby_ATTR :	BYTE;
	END_VAR

	TN_SC_SHADOW_ATTR := ((Iby_ATTR AND BYTE#2#11110000) OR BYTE#2#00001000);

END_FUNCTION

PROGRAM program0
	VAR
		Iby_ATTR :	BYTE;
		CEIL5_OUT : BYTE;
	END_VAR

  	CEIL5_OUT := TN_SC_SHADOW_ATTR(Iby_ATTR);
END_PROGRAM

CONFIGURATION Config0

  RESOURCE Res0 ON PLC
    TASK task0(INTERVAL := T#20ms,PRIORITY := 0);
    PROGRAM instance0 WITH task0 : program0;
  END_RESOURCE
END_CONFIGURATION

(* ---- TN_SC_XY2_ERROR.ST ---- *)
FUNCTION TN_SC_XY2_ERROR:BOOL

	VAR_INPUT
		X1 :	INT;
		Y1 :	INT;
		X2 :	INT;
		Y2 :	INT;
	END_VAR

	TN_SC_XY2_ERROR := Y1 < 0 OR X1 < 0 OR Y2 < 0 OR X2 < 0 OR Y1 > 23 OR X1 > 79 OR Y2 > 23 OR X2 > 79;

END_FUNCTION

PROGRAM program0
	VAR
		X1 :	INT;
		Y1 :	INT;
		X2 :	INT;
		Y2 :	INT;
		CEIL5_OUT : BOOL;
	END_VAR

  	CEIL5_OUT := TN_SC_XY2_ERROR(X1, Y1, X2, Y2);
END_PROGRAM

CONFIGURATION Config0

  RESOURCE Res0 ON PLC
    TASK task0(INTERVAL := T#20ms,PRIORITY := 0);
    PROGRAM instance0 WITH task0 : program0;
  END_RESOURCE
END_CONFIGURATION

(* ---- TN_SC_XY_ERROR.ST ---- *)
FUNCTION TN_SC_XY_ERROR:BOOL

	VAR_INPUT
		X :	INT;
		Y :	INT;
	END_VAR

	TN_SC_XY_ERROR := Y < 0 OR X < 0 OR Y > 23 OR X > 79;

END_FUNCTION

PROGRAM program0
	VAR
		X :	INT;
		Y :	INT;
		CEIL5_OUT : BOOL;
	END_VAR

  	CEIL5_OUT := TN_SC_XY_ERROR(X, Y);
END_PROGRAM

CONFIGURATION Config0

  RESOURCE Res0 ON PLC
    TASK task0(INTERVAL := T#20ms,PRIORITY := 0);
    PROGRAM instance0 WITH task0 : program0;
  END_RESOURCE
END_CONFIGURATION

(* ---- TO_LOWER.ST ---- *)
FUNCTION SETUP_EXTENDED_ASCII:BOOL

	VAR_INPUT
		X :	BOOL;
	END_VAR

	SETUP_EXTENDED_ASCII := X OR TRUE;
END_FUNCTION

FUNCTION TO_LOWER:BYTE

	VAR_INPUT
		IN :	BYTE;
	END_VAR

	IF in > BYTE#64 AND in < BYTE#91 THEN
	TO_LOWER := in OR BYTE#16#20;
	ELSIF (in > BYTE#191 AND in < BYTE#223) AND in <> BYTE#215 AND SETUP_EXTENDED_ASCII(FALSE) THEN
	TO_LOWER := in OR BYTE#16#20;
	ELSE
	TO_LOWER := in;
	END_IF;

END_FUNCTION

PROGRAM program0
  VAR
	IN :	BYTE;
    CEIL5_OUT : BYTE;
  END_VAR

  CEIL5_OUT := TO_LOWER(IN);
END_PROGRAM

CONFIGURATION Config0

  RESOURCE Res0 ON PLC
    TASK task0(INTERVAL := T#20ms,PRIORITY := 0);
    PROGRAM instance0 WITH task0 : program0;
  END_RESOURCE
END_CONFIGURATION

(* ---- TO_UPPER.ST ---- *)
FUNCTION SETUP_EXTENDED_ASCII:BOOL
	VAR_INPUT
		X :	BOOL;
	END_VAR

	SETUP_EXTENDED_ASCII := X OR TRUE;
END_FUNCTION

FUNCTION TO_UPPER:BYTE

	VAR_INPUT
		IN :	BYTE;
	END_VAR

	IF in > BYTE#96 AND in < BYTE#123 THEN
	TO_UPPER := in AND BYTE#16#DF;
	ELSIF in > BYTE#223 AND in <> BYTE#247 AND in <> BYTE#255 AND SETUP_EXTENDED_ASCII(FALSE) THEN
	TO_UPPER := in AND BYTE#16#DF;
	ELSE
	TO_UPPER := in;
	END_IF;

END_FUNCTION

PROGRAM program0
  VAR
	IN :	BYTE;
    CEIL5_OUT : BYTE;
  END_VAR

  CEIL5_OUT := TO_UPPER(IN);
END_PROGRAM

CONFIGURATION Config0

  RESOURCE Res0 ON PLC
    TASK task0(INTERVAL := T#20ms,PRIORITY := 0);
    PROGRAM instance0 WITH task0 : program0;
  END_RESOURCE
END_CONFIGURATION

(* ---- TOD_TO_REAL.ST ---- *)
FUNCTION TOD_TO_REAL2:REAL
	VAR_INPUT
		IN :	UDINT;
	END_VAR
	TOD_TO_REAL2 := UDINT_TO_REAL(IN);
END_FUNCTION

PROGRAM program0
  VAR
	IN :	UDINT;
    CEIL5_OUT : REAL;
  END_VAR

  CEIL5_OUT := TOD_TO_REAL2(IN);
END_PROGRAM

CONFIGURATION Config0

  RESOURCE Res0 ON PLC
    TASK task0(INTERVAL := T#20ms,PRIORITY := 0);
    PROGRAM instance0 WITH task0 : program0;
  END_RESOURCE
END_CONFIGURATION

(* ---- TOD_TO_TIME.ST ---- *)
FUNCTION TOD_TO_TIME:TIME
	VAR_INPUT
		IN :	UDINT;
	END_VAR

	TOD_TO_TIME := DWORD_TO_TIME(UDINT_TO_DWORD(IN));
END_FUNCTION

PROGRAM program0
  VAR
	IN :	UDINT;
    CEIL5_OUT : TIME;
  END_VAR

  CEIL5_OUT := TOD_TO_TIME(IN);
END_PROGRAM

CONFIGURATION Config0

  RESOURCE Res0 ON PLC
    TASK task0(INTERVAL := T#20ms,PRIORITY := 0);
    PROGRAM instance0 WITH task0 : program0;
  END_RESOURCE
END_CONFIGURATION

(* ---- TRIANGLE_A.ST ---- *)
FUNCTION _REAL_TO_DINT:DINT
  VAR_INPUT
    X :	REAL;
  END_VAR

  IF REAL_TO_DINT(0.5) = DINT#1 THEN
    _REAL_TO_DINT := REAL_TO_DINT(x);
    RETURN;
  END_IF;

  IF X > 0.0 THEN
    _REAL_TO_DINT := REAL_TO_DINT(x+0.5);
  ELSIF X < 0.0 THEN
    _REAL_TO_DINT := REAL_TO_DINT(x-0.5);
  ELSE
    _REAL_TO_DINT := DINT#0;
  END_IF;
END_FUNCTION

FUNCTION FLOOR2:DINT

	VAR_INPUT
		X :	REAL;
	END_VAR

	FLOOR2 := _REAL_TO_DINT(X);
	IF DINT_TO_REAL(FLOOR2) > X THEN
		FLOOR2 := FLOOR2 - DINT#1;
	END_IF;

END_FUNCTION

FUNCTION MODR:REAL

	VAR_INPUT
		IN :	REAL;
		DIVI :	REAL;
	END_VAR

	IF divi = 0.0 THEN
		MODR := 0.0;
	ELSE
		MODR := in - DINT_TO_REAL(FLOOR2(in / divi)) * divi;
	END_IF;

END_FUNCTION

FUNCTION RAD:REAL

	VAR_INPUT
		DEG :	REAL;
	END_VAR

	Rad := modR(0.0174532925199433 * deg , 6.283185307179586476);

END_FUNCTION

FUNCTION TRIANGLE_A:REAL

	VAR_INPUT
		S1 :	REAL;
		A :	REAL;
		S2 :	REAL;
		S3 :	REAL;
	END_VAR

	IF A = 0.0 THEN
		TRIANGLE_A := SQRT((s1+s2+S3) * (s1+s2-S3) * (S2+S3-S1) * (S3+S1-S2)) * 0.25;
	ELSE
		TRIANGLE_A := S1 * S2 * SIN(RAD(A)) * 0.5;
	END_IF;

END_FUNCTION

PROGRAM program0
  VAR
	S1 :	REAL;
	A :	REAL;
	S2 :	REAL;
	S3 :	REAL;
    CEIL5_OUT : REAL;
  END_VAR

  CEIL5_OUT := TRIANGLE_A(S1, A, S2, S3);
END_PROGRAM

CONFIGURATION Config0

  RESOURCE Res0 ON PLC
    TASK task0(INTERVAL := T#20ms,PRIORITY := 0);
    PROGRAM instance0 WITH task0 : program0;
  END_RESOURCE
END_CONFIGURATION

(* ---- TRUNC_REAL.ST ---- *)
FUNCTION TRUNC_REAL:REAL

	VAR_INPUT
		IN :	REAL;
	END_VAR

	TRUNC_REAL := UDINT_TO_REAL(DINT_TO_UDINT(TRUNC(IN)));
END_FUNCTION

PROGRAM program0

	VAR
		IN :	REAL;
		OUT: REAL;
	END_VAR
	OUT := TRUNC_REAL(IN);

END_PROGRAM

CONFIGURATION Config0

	RESOURCE Res0 ON PLC
		TASK task0(INTERVAL := T#20ms,PRIORITY := 0);
		PROGRAM instance0 WITH task0 : program0;
	END_RESOURCE

END_CONFIGURATION

(* ---- TRUNC_UDINT.ST ---- *)
FUNCTION TRUNC_UDINT:UDINT
	VAR_INPUT
		IN :	REAL;
	END_VAR
	TRUNC_UDINT := DINT_TO_UDINT(TRUNC(IN));
END_FUNCTION

PROGRAM program0
	VAR
		LocalVar0 : REAL;
		LocalOUT  : UDINT;
	END_VAR
		LocalOUT := TRUNC_UDINT(LocalVar0);
END_PROGRAM

CONFIGURATION Config0
	RESOURCE Res0 ON PLC
		TASK task0(INTERVAL := T#20ms,PRIORITY := 0);
		PROGRAM instance0 WITH task0 : program0;
	END_RESOURCE
END_CONFIGURATION

(* ---- UDINT_TO_TIME.ST ---- *)
FUNCTION _UDINT_TO_TIME:TIME

	VAR_INPUT
		IN :	UDINT;
	END_VAR

	_UDINT_TO_TIME := DINT_TO_TIME(UDINT_TO_DINT(IN));

END_FUNCTION

PROGRAM program0
  VAR
	  IN :	UDINT;
    CEIL5_OUT : TIME;
  END_VAR

  CEIL5_OUT := _UDINT_TO_TIME(IN);
END_PROGRAM

CONFIGURATION Config0

  RESOURCE Res0 ON PLC
    TASK task0(INTERVAL := T#20ms,PRIORITY := 0);
    PROGRAM instance0 WITH task0 : program0;
  END_RESOURCE
END_CONFIGURATION
